(* IEC 61131-3 sources: plc-st-coding-agent/progress/evidence/f14_v6_public_pilot_20261112/jobs/custom_minimax-m27 (part 2) *)

(* ---- public-medium-03.candidate_02.st ---- *)
FUNCTION_BLOCK FB_MovingAverage
VAR_INPUT
    cyclicExecution : BOOL;
    trigger         : BOOL;
    value           : LREAL;
    windowSize      : INT;
    reset           : BOOL;
END_VAR

VAR_OUTPUT
    average           : LREAL;
    windowSizeReached : BOOL;
    error             : BOOL;
    status            : WORD;
END_VAR

VAR
    dataBuffer       : ARRAY[1..100] OF LREAL;
    currentIndex     : INT := 0;
    sampleCount      : INT := 0;
    sum              : LREAL := 0.0;
    tmp_lastTrigger  : BOOL := FALSE;
    tmp_newSample    : BOOL := FALSE;
    tmp_effectiveWin : INT := 0;
END_VAR

(*
ENGINEERING_CONTRACT
===================
Operation Modes:
- cyclicExecution=TRUE: Update every scan cycle; trigger ignored (PUB002)
- cyclicExecution=FALSE: Rising edge on trigger updates average (PUB003)
- reset=TRUE: Clear all state, outputs to default, status=SUCCESS (PUB004)

Output Retention Policy:
| Output             | Activation         | Retention    | Reset by reset=TRUE |
|--------------------|--------------------|--------------|---------------------|
| average            | Each valid sample  | Hold last    | Yes (→0.0)          |
| windowSizeReached  | sampleCount>=winSz | Hold TRUE    | Yes (→FALSE)        |
| error              | windowSize<1 or >100| Hold TRUE   | Yes (→FALSE)        |
| status             | Per validation     | Hold code    | Yes (→SUCCESS)      |

Boundary Conditions:
- windowSize<1 OR >100 → error=TRUE, status=16#8200, skip processing (PUB004, PUB007)
- reset asserted → immediate clear, no processing (PUB004)
- Empty window (sampleCount=0) → average=0.0 (division-safe)
- Circular buffer wraps at windowSize, never exceeds 100 elements

Same-Scan Priority:
1. reset check (highest)
2. windowSize validation
3. trigger rising-edge detection
4. cyclicExecution evaluation
5. sample insertion / buffer rotation
6. average recalculation

Units: LREAL for all arithmetic (PUB001). windowSize in slots [1..100].
*)

(* CONTRACT_RULES
[
  {"kind": "hold_until_reset", "output": "windowSizeReached", "set_input": null, "reset_input": "reset"},
  {"kind": "hold_until_reset", "output": "error", "set_input": null, "reset_input": "reset"},
  {"kind": "hold_until_reset", "output": "status", "set_input": null, "reset_input": "reset"}
]
*)

    // Reset: clear all state and outputs
    IF reset THEN
        currentIndex      := 0;
        sampleCount       := 0;
        sum               := 0.0;
        average           := 0.0;
        windowSizeReached := FALSE;
        error             := FALSE;
        status            := 16#0000;
        tmp_lastTrigger   := FALSE;
        tmp_newSample     := FALSE;
        tmp_effectiveWin  := 0;
        RETURN;
    END_IF;

    // Validate window size (PUB007)
    IF windowSize < 1 OR windowSize > 100 THEN
        error  := TRUE;
        status := 16#8200;
        RETURN;
    END_IF;

    // No validation error; set success status (PUB006)
    error  := FALSE;
    status := 16#0000;

    // Determine if a new sample should be processed (PUB002, PUB003)
    tmp_newSample := FALSE;
    IF cyclicExecution THEN
        tmp_newSample := TRUE;
    ELSIF trigger AND NOT tmp_lastTrigger THEN
        tmp_newSample := TRUE;
    END_IF;
    tmp_lastTrigger := trigger;

    // Process new data point if triggered (PUB001)
    IF tmp_newSample THEN
        // Clamp effective window to array upper bound (100)
        tmp_effectiveWin := windowSize;
        IF tmp_effectiveWin > 100 THEN
            tmp_effectiveWin := 100;
        END_IF;

        IF sampleCount < tmp_effectiveWin THEN
            // Window not yet full: append new value
            sampleCount := sampleCount + 1;
            dataBuffer[sampleCount] := value;
            sum := sum + value;
        ELSE
            // Window full: rotate out oldest value using circular buffer
            currentIndex := (currentIndex MOD tmp_effectiveWin) + 1;
            sum := sum - dataBuffer[currentIndex] + value;
            dataBuffer[currentIndex] := value;
        END_IF;
    END_IF;

    // Calculate moving arithmetic mean (PUB001)
    IF sampleCount > 0 THEN
        average := sum / TO_LREAL(sampleCount);
    ELSE
        average := 0.0;
    END_IF;

    // Indicate whether maximum window width has been reached (PUB001)
    tmp_effectiveWin := windowSize;
    IF tmp_effectiveWin > 100 THEN
        tmp_effectiveWin := 100;
    END_IF;
    windowSizeReached := (sampleCount >= tmp_effectiveWin);

END_FUNCTION_BLOCK

(* ---- public-medium-03.candidate_03.st ---- *)
FUNCTION_BLOCK FB_MovingAverage
VAR_INPUT
    cyclicExecution : BOOL;
    trigger         : BOOL;
    value           : LREAL;
    windowSize      : INT;
    reset           : BOOL;
END_VAR

VAR_OUTPUT
    average           : LREAL;
    windowSizeReached : BOOL;
    error             : BOOL;
    status            : WORD;
END_VAR

VAR
    dataBuffer       : ARRAY[1..100] OF LREAL;
    sampleCount      : INT := 0;
    sum              : LREAL := 0.0;
    tmp_lastTrigger  : BOOL := FALSE;
    tmp_effectiveWin : INT := 0;
END_VAR

(*
ENGINEERING_CONTRACT
===================
Operation Modes:
- cyclicExecution=TRUE: Update every scan cycle; trigger ignored (PUB002)
- cyclicExecution=FALSE: Rising edge on trigger updates average (PUB003)
- reset=TRUE: Clear all state, outputs to default, status=SUCCESS (PUB004)

Output Retention Policy:
| Output             | Activation         | Retention    | Reset by reset=TRUE |
|--------------------|--------------------|--------------|---------------------|
| average            | Each valid sample  | Hold last    | Yes (→0.0)          |
| windowSizeReached  | sampleCount>=winSz | Hold TRUE    | Yes (→FALSE)        |
| error              | windowSize<1 or >100| Hold TRUE   | Yes (→FALSE)        |
| status             | Per validation     | Hold code    | Yes (→SUCCESS)      |

Boundary Conditions:
- windowSize<1 OR >100 → error=TRUE, status=16#8200, skip processing (PUB004, PUB007)
- reset asserted → immediate clear, no processing (PUB004)
- Empty window (sampleCount=0) → average=0.0 (division-safe)
- Circular buffer wraps at windowSize, never exceeds 100 elements

Same-Scan Priority:
1. reset check (highest)
2. windowSize validation
3. trigger rising-edge detection
4. cyclicExecution evaluation
5. sample insertion / buffer rotation
6. average recalculation

Units: LREAL for all arithmetic (PUB001). windowSize in slots [1..100].
*)

(* CONTRACT_RULES
[
  {"kind": "hold_until_reset", "output": "windowSizeReached", "set_input": null, "reset_input": "reset"},
  {"kind": "hold_until_reset", "output": "error", "set_input": null, "reset_input": "reset"},
  {"kind": "hold_until_reset", "output": "status", "set_input": null, "reset_input": "reset"}
]
*)

    // Reset: clear all state and outputs
    IF reset THEN
        sampleCount       := 0;
        sum               := 0.0;
        average           := 0.0;
        windowSizeReached := FALSE;
        error             := FALSE;
        status            := 16#0000;
        tmp_lastTrigger   := FALSE;
        tmp_effectiveWin  := 0;
        RETURN;
    END_IF;

    // Validate window size (PUB007)
    IF windowSize < 1 OR windowSize > 100 THEN
        error  := TRUE;
        status := 16#8200;
        RETURN;
    END_IF;

    // No validation error; set success status (PUB006)
    error  := FALSE;
    status := 16#0000;

    // Clamp effective window to array upper bound (100)
    tmp_effectiveWin := windowSize;
    IF tmp_effectiveWin > 100 THEN
        tmp_effectiveWin := 100;
    END_IF;

    // Determine if a new sample should be processed (PUB002, PUB003)
    IF cyclicExecution OR (trigger AND NOT tmp_lastTrigger) THEN
        // Process new data point (PUB001)
        IF sampleCount < tmp_effectiveWin THEN
            // Window not yet full: append new value
            sampleCount := sampleCount + 1;
            dataBuffer[sampleCount] := value;
            sum := sum + value;
        ELSE
            // Window full: rotate out oldest value
            // Shift all elements down by one position
            sum := sum - dataBuffer[1];
            FOR i := 1 TO tmp_effectiveWin - 1 DO
                dataBuffer[i] := dataBuffer[i + 1];
            END_FOR;
            dataBuffer[tmp_effectiveWin] := value;
            sum := sum + value;
        END_IF;
    END_IF;

    // Update trigger state for edge detection
    tmp_lastTrigger := trigger;

    // Calculate moving arithmetic mean (PUB001)
    IF sampleCount > 0 THEN
        average := sum / TO_LREAL(sampleCount);
    ELSE
        average := 0.0;
    END_IF;

    // Indicate whether maximum window width has been reached (PUB001)
    windowSizeReached := (sampleCount >= tmp_effectiveWin);

END_FUNCTION_BLOCK

(* ---- public-medium-03.candidate_04.st ---- *)
FUNCTION_BLOCK FB_MovingAverage
VAR_INPUT
    cyclicExecution : BOOL;
    trigger         : BOOL;
    value           : LREAL;
    windowSize      : INT;
    reset           : BOOL;
END_VAR

VAR_OUTPUT
    average           : LREAL;
    windowSizeReached : BOOL;
    error             : BOOL;
    status            : WORD;
END_VAR

VAR
    dataBuffer         : ARRAY[1..100] OF LREAL;
    currentIndex       : INT := 0;
    sampleCount        : INT := 0;
    sum                : LREAL := 0.0;
    tmp_lastTrigger    : BOOL := FALSE;
    tmp_newSample      : BOOL := FALSE;
    tmp_effectiveWin   : INT := 0;
    tmp_winSizeChanged : BOOL := FALSE;
    tmp_prevWinSize    : INT := 0;
    tmp_startIdx       : INT := 0;
    tmp_i              : INT := 0;
    tmp_newSum         : LREAL := 0.0;
END_VAR

(*
ENGINEERING_CONTRACT
===================
Operation Modes:
- cyclicExecution=TRUE: Update every scan cycle; trigger ignored (PUB002)
- cyclicExecution=FALSE: Rising edge on trigger updates average (PUB003)
- reset=TRUE: Clear all state, outputs to default, status=SUCCESS (PUB004)

Output Retention Policy:
| Output             | Activation         | Retention    | Reset by reset=TRUE |
|--------------------|--------------------|--------------|---------------------|
| average            | Each valid sample  | Hold last    | Yes (→0.0)          |
| windowSizeReached  | sampleCount>=winSz | Hold TRUE    | Yes (→FALSE)        |
| error              | windowSize<1 or >100| Hold TRUE   | Yes (→FALSE)        |
| status             | Per validation     | Hold code    | Yes (→SUCCESS)      |

Boundary Conditions:
- windowSize<1 OR >100 → error=TRUE, status=16#8200, skip processing (PUB004, PUB007)
- reset asserted → immediate clear, no processing (PUB004)
- Empty window (sampleCount=0) → average=0.0 (division-safe)
- Circular buffer wraps at windowSize, never exceeds 100 elements
- windowSize change → prune buffer to contain only most recent windowSize samples

Same-Scan Priority:
1. reset check (highest)
2. windowSize validation (set error=TRUE if invalid, return)
3. windowSize change detection → prune buffer
4. trigger rising-edge detection
5. cyclicExecution evaluation
6. sample insertion / buffer rotation
7. average recalculation

Units: LREAL for all arithmetic (PUB001). windowSize in slots [1..100].
*)

(* CONTRACT_RULES
[
  {"kind": "hold_until_reset", "output": "windowSizeReached", "set_input": null, "reset_input": "reset"},
  {"kind": "hold_until_reset", "output": "error", "set_input": null, "reset_input": "reset"},
  {"kind": "hold_until_reset", "output": "status", "set_input": null, "reset_input": "reset"}
]
*)

    // Reset: clear all state and outputs
    IF reset THEN
        currentIndex      := 0;
        sampleCount       := 0;
        sum               := 0.0;
        average           := 0.0;
        windowSizeReached := FALSE;
        error             := FALSE;
        status            := 16#0000;
        tmp_lastTrigger   := FALSE;
        tmp_newSample     := FALSE;
        tmp_effectiveWin  := 0;
        tmp_winSizeChanged := FALSE;
        tmp_prevWinSize   := 0;
        tmp_startIdx      := 0;
        tmp_i             := 0;
        tmp_newSum        := 0.0;
        RETURN;
    END_IF;

    // Clamp effective window to array upper bound for validation
    tmp_effectiveWin := windowSize;
    IF tmp_effectiveWin > 100 THEN
        tmp_effectiveWin := 100;
    END_IF;

    // Validate window size (PUB007)
    // Only clear error AFTER validation passes, so invalid sizes preserve error state
    IF windowSize < 1 OR windowSize > 100 THEN
        error  := TRUE;
        status := 16#8200;
        RETURN;
    END_IF;

    // Valid windowSize: clear error and set success status (PUB006)
    error  := FALSE;
    status := 16#0000;

    // Detect windowSize change and prune buffer if needed
    tmp_winSizeChanged := (tmp_prevWinSize <> 0) AND (tmp_prevWinSize <> windowSize);
    IF tmp_winSizeChanged AND sampleCount > 0 THEN
        // Prune buffer to contain only most recent windowSize samples
        tmp_effectiveWin := windowSize;
        IF tmp_effectiveWin > 100 THEN
            tmp_effectiveWin := 100;
        END_IF;

        IF sampleCount > tmp_effectiveWin THEN
            // Calculate start index for circular buffer (oldest sample to keep)
            // Most recent samples are at positions (currentIndex - k + 1) through currentIndex
            tmp_startIdx := ((currentIndex - tmp_effectiveWin) MOD 100) + 1;
            IF tmp_startIdx < 1 THEN
                tmp_startIdx := tmp_startIdx + 100;
            END_IF;

            // Copy most recent samples to front of buffer and recalculate sum
            tmp_newSum := 0.0;
            FOR tmp_i := 1 TO tmp_effectiveWin DO
                dataBuffer[tmp_i] := dataBuffer[tmp_startIdx + tmp_i - 1];
                tmp_newSum := tmp_newSum + dataBuffer[tmp_i];
            END_FOR;

            // Clear remaining buffer slots
            FOR tmp_i := tmp_effectiveWin + 1 TO 100 DO
                dataBuffer[tmp_i] := 0.0;
            END_FOR;

            sampleCount := tmp_effectiveWin;
            sum := tmp_newSum;
            currentIndex := tmp_effectiveWin;
        END_IF;
    END_IF;

    // Track current windowSize for next-cycle change detection
    tmp_prevWinSize := windowSize;

    // Determine if a new sample should be processed (PUB002, PUB003)
    tmp_newSample := FALSE;
    IF cyclicExecution THEN
        tmp_newSample := TRUE;
    ELSIF trigger AND NOT tmp_lastTrigger THEN
        tmp_newSample := TRUE;
    END_IF;
    tmp_lastTrigger := trigger;

    // Process new data point if triggered (PUB001)
    IF tmp_newSample THEN
        tmp_effectiveWin := windowSize;
        IF tmp_effectiveWin > 100 THEN
            tmp_effectiveWin := 100;
        END_IF;

        IF sampleCount < tmp_effectiveWin THEN
            // Buffer not yet full: append new value
            sampleCount := sampleCount + 1;
            currentIndex := sampleCount;
            dataBuffer[currentIndex] := value;
            sum := sum + value;
        ELSE
            // Buffer full: rotate out oldest value using circular buffer
            currentIndex := (currentIndex MOD tmp_effectiveWin) + 1;
            sum := sum - dataBuffer[currentIndex] + value;
            dataBuffer[currentIndex] := value;
        END_IF;
    END_IF;

    // Calculate moving arithmetic mean (PUB001)
    IF sampleCount > 0 THEN
        average := sum / TO_LREAL(sampleCount);
    ELSE
        average := 0.0;
    END_IF;

    // Indicate whether maximum window width has been reached (PUB001)
    tmp_effectiveWin := windowSize;
    IF tmp_effectiveWin > 100 THEN
        tmp_effectiveWin := 100;
    END_IF;
    windowSizeReached := (sampleCount >= tmp_effectiveWin);

END_FUNCTION_BLOCK

(* ---- public-medium-03.raw_candidate_01.st ---- *)
FUNCTION_BLOCK FB_MovingAverage
VAR_INPUT
    cyclicExecution : BOOL;
    trigger         : BOOL;
    value           : LREAL;
    windowSize      : INT;
    reset           : BOOL;
END_VAR

VAR_OUTPUT
    average           : LREAL;
    windowSizeReached : BOOL;
    error             : BOOL;
    status            : WORD;
END_VAR

VAR
    dataBuffer    : ARRAY[1..100] OF LREAL;
    currentIndex  : INT := 0;
    sampleCount   : INT := 0;
    sum           : LREAL := 0.0;
    tmp_lastTrigger : BOOL := FALSE;
END_VAR

(*
ENGINEERING_CONTRACT
===================
Operation Modes:
- cyclicExecution=TRUE: Update every scan cycle; trigger ignored (PUB002)
- cyclicExecution=FALSE: Rising edge on trigger updates average (PUB003)
- reset=TRUE: Clear all state, outputs to default, status=SUCCESS (PUB004)

Output Retention Policy:
| Output             | Activation         | Retention    | Reset by reset=TRUE |
|--------------------|--------------------|--------------|---------------------|
| average            | Each valid sample  | Hold last    | Yes (→0.0)          |
| windowSizeReached  | sampleCount>=winSz | Hold TRUE    | Yes (→FALSE)        |
| error              | windowSize<1 or >100| Hold TRUE   | Yes (→FALSE)        |
| status             | Per validation     | Hold code    | Yes (→SUCCESS)      |

Boundary Conditions:
- windowSize<1 OR >100 → error=TRUE, status=16#8200, skip processing (PUB004, PUB007)
- reset asserted → immediate clear, no processing (PUB004)
- Empty window (sampleCount=0) → average=0.0 (division-safe)
- Circular buffer wraps at windowSize, never exceeds 100 elements

Same-Scan Priority:
1. reset check (highest)
2. windowSize validation
3. trigger rising-edge detection
4. cyclicExecution evaluation
5. sample insertion / buffer rotation
6. average recalculation

Units: LREAL for all arithmetic (PUB001). windowSize in slots [1..100].
*)

(* CONTRACT_RULES
[
  {"kind": "hold_until_reset", "output": "windowSizeReached", "set_input": null, "reset_input": "reset"},
  {"kind": "hold_until_reset", "output": "error", "set_input": null, "reset_input": "reset"},
  {"kind": "hold_until_reset", "output": "status", "set_input": null, "reset_input": "reset"}
]
*)

    // Reset: clear all state and outputs
    IF reset THEN
        currentIndex     := 0;
        sampleCount      := 0;
        sum              := 0.0;
        average          := 0.0;
        windowSizeReached := FALSE;
        error            := FALSE;
        status           := 16#0000;
        tmp_lastTrigger  := FALSE;
        RETURN;
    END_IF

    // Validate window size (PUB007)
    IF windowSize < 1 OR windowSize > 100 THEN
        error  := TRUE;
        status := 16#8200;
        RETURN;
    END_IF

    // No validation error; set success status (PUB006)
    error  := FALSE;
    status := 16#0000;

    // Determine if a new sample should be processed (PUB002, PUB003)
    tmp_newSample := FALSE;
    IF cyclicExecution THEN
        tmp_newSample := TRUE;
    ELSIF trigger AND NOT tmp_lastTrigger THEN
        tmp_newSample := TRUE;
    END_IF
    tmp_lastTrigger := trigger;

    // Process new data point if triggered (PUB001)
    IF tmp_newSample THEN
        // Clamp effective window to array upper bound (100)
        tmp_effectiveWindow := windowSize;
        IF tmp_effectiveWindow > 100 THEN
            tmp_effectiveWindow := 100;
        END_IF

        IF sampleCount < tmp_effectiveWindow THEN
            // Window not yet full: append new value
            sampleCount := sampleCount + 1;
            dataBuffer[sampleCount] := value;
            sum := sum + value;
        ELSE
            // Window full: rotate out oldest value using circular buffer
            currentIndex := (currentIndex MOD tmp_effectiveWindow) + 1;
            sum := sum - dataBuffer[currentIndex] + value;
            dataBuffer[currentIndex] := value;
        END_IF
    END_IF

    // Calculate moving arithmetic mean (PUB001)
    IF sampleCount > 0 THEN
        average := sum / TO_LREAL(sampleCount);
    ELSE
        average := 0.0;
    END_IF

    // Indicate whether maximum window width has been reached (PUB001)
    tmp_effectiveWindow := windowSize;
    IF tmp_effectiveWindow > 100 THEN
        tmp_effectiveWindow := 100;
    END_IF;
    windowSizeReached := (sampleCount >= tmp_effectiveWindow);

END_FUNCTION_BLOCK

(* ---- public-medium-03.raw_candidate_02.st ---- *)
FUNCTION_BLOCK FB_MovingAverage
VAR_INPUT
    cyclicExecution : BOOL;
    trigger         : BOOL;
    value           : LREAL;
    windowSize      : INT;
    reset           : BOOL;
END_VAR

VAR_OUTPUT
    average           : LREAL;
    windowSizeReached : BOOL;
    error             : BOOL;
    status            : WORD;
END_VAR

VAR
    dataBuffer       : ARRAY[1..100] OF LREAL;
    currentIndex     : INT := 0;
    sampleCount      : INT := 0;
    sum              : LREAL := 0.0;
    tmp_lastTrigger  : BOOL := FALSE;
    tmp_newSample    : BOOL := FALSE;
    tmp_effectiveWin : INT := 0;
END_VAR

(*
ENGINEERING_CONTRACT
===================
Operation Modes:
- cyclicExecution=TRUE: Update every scan cycle; trigger ignored (PUB002)
- cyclicExecution=FALSE: Rising edge on trigger updates average (PUB003)
- reset=TRUE: Clear all state, outputs to default, status=SUCCESS (PUB004)

Output Retention Policy:
| Output             | Activation         | Retention    | Reset by reset=TRUE |
|--------------------|--------------------|--------------|---------------------|
| average            | Each valid sample  | Hold last    | Yes (→0.0)          |
| windowSizeReached  | sampleCount>=winSz | Hold TRUE    | Yes (→FALSE)        |
| error              | windowSize<1 or >100| Hold TRUE   | Yes (→FALSE)        |
| status             | Per validation     | Hold code    | Yes (→SUCCESS)      |

Boundary Conditions:
- windowSize<1 OR >100 → error=TRUE, status=16#8200, skip processing (PUB004, PUB007)
- reset asserted → immediate clear, no processing (PUB004)
- Empty window (sampleCount=0) → average=0.0 (division-safe)
- Circular buffer wraps at windowSize, never exceeds 100 elements

Same-Scan Priority:
1. reset check (highest)
2. windowSize validation
3. trigger rising-edge detection
4. cyclicExecution evaluation
5. sample insertion / buffer rotation
6. average recalculation

Units: LREAL for all arithmetic (PUB001). windowSize in slots [1..100].
*)

(* CONTRACT_RULES
[
  {"kind": "hold_until_reset", "output": "windowSizeReached", "set_input": null, "reset_input": "reset"},
  {"kind": "hold_until_reset", "output": "error", "set_input": null, "reset_input": "reset"},
  {"kind": "hold_until_reset", "output": "status", "set_input": null, "reset_input": "reset"}
]
*)

    // Reset: clear all state and outputs
    IF reset THEN
        currentIndex      := 0;
        sampleCount       := 0;
        sum               := 0.0;
        average           := 0.0;
        windowSizeReached := FALSE;
        error             := FALSE;
        status            := 16#0000;
        tmp_lastTrigger   := FALSE;
        tmp_newSample     := FALSE;
        tmp_effectiveWin  := 0;
        RETURN;
    END_IF;

    // Validate window size (PUB007)
    IF windowSize < 1 OR windowSize > 100 THEN
        error  := TRUE;
        status := 16#8200;
        RETURN;
    END_IF;

    // No validation error; set success status (PUB006)
    error  := FALSE;
    status := 16#0000;

    // Determine if a new sample should be processed (PUB002, PUB003)
    tmp_newSample := FALSE;
    IF cyclicExecution THEN
        tmp_newSample := TRUE;
    ELSIF trigger AND NOT tmp_lastTrigger THEN
        tmp_newSample := TRUE;
    END_IF;
    tmp_lastTrigger := trigger;

    // Process new data point if triggered (PUB001)
    IF tmp_newSample THEN
        // Clamp effective window to array upper bound (100)
        tmp_effectiveWin := windowSize;
        IF tmp_effectiveWin > 100 THEN
            tmp_effectiveWin := 100;
        END_IF;

        IF sampleCount < tmp_effectiveWin THEN
            // Window not yet full: append new value
            sampleCount := sampleCount + 1;
            dataBuffer[sampleCount] := value;
            sum := sum + value;
        ELSE
            // Window full: rotate out oldest value using circular buffer
            currentIndex := (currentIndex MOD tmp_effectiveWin) + 1;
            sum := sum - dataBuffer[currentIndex] + value;
            dataBuffer[currentIndex] := value;
        END_IF;
    END_IF;

    // Calculate moving arithmetic mean (PUB001)
    IF sampleCount > 0 THEN
        average := sum / TO_LREAL(sampleCount);
    ELSE
        average := 0.0;
    END_IF;

    // Indicate whether maximum window width has been reached (PUB001)
    tmp_effectiveWin := windowSize;
    IF tmp_effectiveWin > 100 THEN
        tmp_effectiveWin := 100;
    END_IF;
    windowSizeReached := (sampleCount >= tmp_effectiveWin);

END_FUNCTION_BLOCK

(* ---- public-medium-03.raw_candidate_03.st ---- *)
FUNCTION_BLOCK FB_MovingAverage
VAR_INPUT
    cyclicExecution : BOOL;
    trigger         : BOOL;
    value           : LREAL;
    windowSize      : INT;
    reset           : BOOL;
END_VAR

VAR_OUTPUT
    average           : LREAL;
    windowSizeReached : BOOL;
    error             : BOOL;
    status            : WORD;
END_VAR

VAR
    dataBuffer       : ARRAY[1..100] OF LREAL;
    sampleCount      : INT := 0;
    sum              : LREAL := 0.0;
    tmp_lastTrigger  : BOOL := FALSE;
    tmp_effectiveWin : INT := 0;
END_VAR

(*
ENGINEERING_CONTRACT
===================
Operation Modes:
- cyclicExecution=TRUE: Update every scan cycle; trigger ignored (PUB002)
- cyclicExecution=FALSE: Rising edge on trigger updates average (PUB003)
- reset=TRUE: Clear all state, outputs to default, status=SUCCESS (PUB004)

Output Retention Policy:
| Output             | Activation         | Retention    | Reset by reset=TRUE |
|--------------------|--------------------|--------------|---------------------|
| average            | Each valid sample  | Hold last    | Yes (→0.0)          |
| windowSizeReached  | sampleCount>=winSz | Hold TRUE    | Yes (→FALSE)        |
| error              | windowSize<1 or >100| Hold TRUE   | Yes (→FALSE)        |
| status             | Per validation     | Hold code    | Yes (→SUCCESS)      |

Boundary Conditions:
- windowSize<1 OR >100 → error=TRUE, status=16#8200, skip processing (PUB004, PUB007)
- reset asserted → immediate clear, no processing (PUB004)
- Empty window (sampleCount=0) → average=0.0 (division-safe)
- Circular buffer wraps at windowSize, never exceeds 100 elements

Same-Scan Priority:
1. reset check (highest)
2. windowSize validation
3. trigger rising-edge detection
4. cyclicExecution evaluation
5. sample insertion / buffer rotation
6. average recalculation

Units: LREAL for all arithmetic (PUB001). windowSize in slots [1..100].
*)

(* CONTRACT_RULES
[
  {"kind": "hold_until_reset", "output": "windowSizeReached", "set_input": null, "reset_input": "reset"},
  {"kind": "hold_until_reset", "output": "error", "set_input": null, "reset_input": "reset"},
  {"kind": "hold_until_reset", "output": "status", "set_input": null, "reset_input": "reset"}
]
*)

    // Reset: clear all state and outputs
    IF reset THEN
        sampleCount       := 0;
        sum               := 0.0;
        average           := 0.0;
        windowSizeReached := FALSE;
        error             := FALSE;
        status            := 16#0000;
        tmp_lastTrigger   := FALSE;
        tmp_effectiveWin  := 0;
        RETURN;
    END_IF;

    // Validate window size (PUB007)
    IF windowSize < 1 OR windowSize > 100 THEN
        error  := TRUE;
        status := 16#8200;
        RETURN;
    END_IF;

    // No validation error; set success status (PUB006)
    error  := FALSE;
    status := 16#0000;

    // Clamp effective window to array upper bound (100)
    tmp_effectiveWin := windowSize;
    IF tmp_effectiveWin > 100 THEN
        tmp_effectiveWin := 100;
    END_IF;

    // Determine if a new sample should be processed (PUB002, PUB003)
    IF cyclicExecution OR (trigger AND NOT tmp_lastTrigger) THEN
        // Process new data point (PUB001)
        IF sampleCount < tmp_effectiveWin THEN
            // Window not yet full: append new value
            sampleCount := sampleCount + 1;
            dataBuffer[sampleCount] := value;
            sum := sum + value;
        ELSE
            // Window full: rotate out oldest value
            // Shift all elements down by one position
            sum := sum - dataBuffer[1];
            FOR i := 1 TO tmp_effectiveWin - 1 DO
                dataBuffer[i] := dataBuffer[i + 1];
            END_FOR;
            dataBuffer[tmp_effectiveWin] := value;
            sum := sum + value;
        END_IF;
    END_IF;

    // Update trigger state for edge detection
    tmp_lastTrigger := trigger;

    // Calculate moving arithmetic mean (PUB001)
    IF sampleCount > 0 THEN
        average := sum / TO_LREAL(sampleCount);
    ELSE
        average := 0.0;
    END_IF;

    // Indicate whether maximum window width has been reached (PUB001)
    windowSizeReached := (sampleCount >= tmp_effectiveWin);

END_FUNCTION_BLOCK

(* ---- public-medium-03.raw_candidate_04.st ---- *)
FUNCTION_BLOCK FB_MovingAverage
VAR_INPUT
    cyclicExecution : BOOL;
    trigger         : BOOL;
    value           : LREAL;
    windowSize      : INT;
    reset           : BOOL;
END_VAR

VAR_OUTPUT
    average           : LREAL;
    windowSizeReached : BOOL;
    error             : BOOL;
    status            : WORD;
END_VAR

VAR
    dataBuffer         : ARRAY[1..100] OF LREAL;
    currentIndex       : INT := 0;
    sampleCount        : INT := 0;
    sum                : LREAL := 0.0;
    tmp_lastTrigger    : BOOL := FALSE;
    tmp_newSample      : BOOL := FALSE;
    tmp_effectiveWin   : INT := 0;
    tmp_winSizeChanged : BOOL := FALSE;
    tmp_prevWinSize    : INT := 0;
    tmp_startIdx       : INT := 0;
    tmp_i              : INT := 0;
    tmp_newSum         : LREAL := 0.0;
END_VAR

(*
ENGINEERING_CONTRACT
===================
Operation Modes:
- cyclicExecution=TRUE: Update every scan cycle; trigger ignored (PUB002)
- cyclicExecution=FALSE: Rising edge on trigger updates average (PUB003)
- reset=TRUE: Clear all state, outputs to default, status=SUCCESS (PUB004)

Output Retention Policy:
| Output             | Activation         | Retention    | Reset by reset=TRUE |
|--------------------|--------------------|--------------|---------------------|
| average            | Each valid sample  | Hold last    | Yes (→0.0)          |
| windowSizeReached  | sampleCount>=winSz | Hold TRUE    | Yes (→FALSE)        |
| error              | windowSize<1 or >100| Hold TRUE   | Yes (→FALSE)        |
| status             | Per validation     | Hold code    | Yes (→SUCCESS)      |

Boundary Conditions:
- windowSize<1 OR >100 → error=TRUE, status=16#8200, skip processing (PUB004, PUB007)
- reset asserted → immediate clear, no processing (PUB004)
- Empty window (sampleCount=0) → average=0.0 (division-safe)
- Circular buffer wraps at windowSize, never exceeds 100 elements
- windowSize change → prune buffer to contain only most recent windowSize samples

Same-Scan Priority:
1. reset check (highest)
2. windowSize validation (set error=TRUE if invalid, return)
3. windowSize change detection → prune buffer
4. trigger rising-edge detection
5. cyclicExecution evaluation
6. sample insertion / buffer rotation
7. average recalculation

Units: LREAL for all arithmetic (PUB001). windowSize in slots [1..100].
*)

(* CONTRACT_RULES
[
  {"kind": "hold_until_reset", "output": "windowSizeReached", "set_input": null, "reset_input": "reset"},
  {"kind": "hold_until_reset", "output": "error", "set_input": null, "reset_input": "reset"},
  {"kind": "hold_until_reset", "output": "status", "set_input": null, "reset_input": "reset"}
]
*)

    // Reset: clear all state and outputs
    IF reset THEN
        currentIndex      := 0;
        sampleCount       := 0;
        sum               := 0.0;
        average           := 0.0;
        windowSizeReached := FALSE;
        error             := FALSE;
        status            := 16#0000;
        tmp_lastTrigger   := FALSE;
        tmp_newSample     := FALSE;
        tmp_effectiveWin  := 0;
        tmp_winSizeChanged := FALSE;
        tmp_prevWinSize   := 0;
        tmp_startIdx      := 0;
        tmp_i             := 0;
        tmp_newSum        := 0.0;
        RETURN;
    END_IF;

    // Clamp effective window to array upper bound for validation
    tmp_effectiveWin := windowSize;
    IF tmp_effectiveWin > 100 THEN
        tmp_effectiveWin := 100;
    END_IF;

    // Validate window size (PUB007)
    // Only clear error AFTER validation passes, so invalid sizes preserve error state
    IF windowSize < 1 OR windowSize > 100 THEN
        error  := TRUE;
        status := 16#8200;
        RETURN;
    END_IF;

    // Valid windowSize: clear error and set success status (PUB006)
    error  := FALSE;
    status := 16#0000;

    // Detect windowSize change and prune buffer if needed
    tmp_winSizeChanged := (tmp_prevWinSize <> 0) AND (tmp_prevWinSize <> windowSize);
    IF tmp_winSizeChanged AND sampleCount > 0 THEN
        // Prune buffer to contain only most recent windowSize samples
        tmp_effectiveWin := windowSize;
        IF tmp_effectiveWin > 100 THEN
            tmp_effectiveWin := 100;
        END_IF;

        IF sampleCount > tmp_effectiveWin THEN
            // Calculate start index for circular buffer (oldest sample to keep)
            // Most recent samples are at positions (currentIndex - k + 1) through currentIndex
            tmp_startIdx := ((currentIndex - tmp_effectiveWin) MOD 100) + 1;
            IF tmp_startIdx < 1 THEN
                tmp_startIdx := tmp_startIdx + 100;
            END_IF;

            // Copy most recent samples to front of buffer and recalculate sum
            tmp_newSum := 0.0;
            FOR tmp_i := 1 TO tmp_effectiveWin DO
                dataBuffer[tmp_i] := dataBuffer[tmp_startIdx + tmp_i - 1];
                tmp_newSum := tmp_newSum + dataBuffer[tmp_i];
            END_FOR;

            // Clear remaining buffer slots
            FOR tmp_i := tmp_effectiveWin + 1 TO 100 DO
                dataBuffer[tmp_i] := 0.0;
            END_FOR;

            sampleCount := tmp_effectiveWin;
            sum := tmp_newSum;
            currentIndex := tmp_effectiveWin;
        END_IF;
    END_IF;

    // Track current windowSize for next-cycle change detection
    tmp_prevWinSize := windowSize;

    // Determine if a new sample should be processed (PUB002, PUB003)
    tmp_newSample := FALSE;
    IF cyclicExecution THEN
        tmp_newSample := TRUE;
    ELSIF trigger AND NOT tmp_lastTrigger THEN
        tmp_newSample := TRUE;
    END_IF;
    tmp_lastTrigger := trigger;

    // Process new data point if triggered (PUB001)
    IF tmp_newSample THEN
        tmp_effectiveWin := windowSize;
        IF tmp_effectiveWin > 100 THEN
            tmp_effectiveWin := 100;
        END_IF;

        IF sampleCount < tmp_effectiveWin THEN
            // Buffer not yet full: append new value
            sampleCount := sampleCount + 1;
            currentIndex := sampleCount;
            dataBuffer[currentIndex] := value;
            sum := sum + value;
        ELSE
            // Buffer full: rotate out oldest value using circular buffer
            currentIndex := (currentIndex MOD tmp_effectiveWin) + 1;
            sum := sum - dataBuffer[currentIndex] + value;
            dataBuffer[currentIndex] := value;
        END_IF;
    END_IF;

    // Calculate moving arithmetic mean (PUB001)
    IF sampleCount > 0 THEN
        average := sum / TO_LREAL(sampleCount);
    ELSE
        average := 0.0;
    END_IF;

    // Indicate whether maximum window width has been reached (PUB001)
    tmp_effectiveWin := windowSize;
    IF tmp_effectiveWin > 100 THEN
        tmp_effectiveWin := 100;
    END_IF;
    windowSizeReached := (sampleCount >= tmp_effectiveWin);

END_FUNCTION_BLOCK

(* ---- public-medium-04.candidate_01.st ---- *)
FUNCTION_BLOCK FBTemperatureControl
VAR_INPUT
    TemperatureSensorInput : REAL;
    SetTemperature         : REAL;
END_VAR
VAR_OUTPUT
    CurrentTemperature : REAL;
    SetTempDisplay     : REAL;
    HeaterStatus       : BOOL;
    OverheatProtection : BOOL;
    HeaterOutput       : BOOL := FALSE;
END_VAR
VAR
    tonHeaterRuntime   : TON;
    tonOverheatCooldown: TON;
    tmpSensorFault     : BOOL;
    tmpHeaterShouldBeOn: BOOL;
END_VAR

(* ENGINEERING_CONTRACT:
 * | State/Output       | Activation                          | Retention           | Reset/Deactivation                                      | Same-scan Priority     | Units/Boundaries   |
 * |--------------------|-------------------------------------|---------------------|---------------------------------------------------------|------------------------|--------------------|
 * | HeaterOutput       | Temp < SetTemp AND no fault AND no overheat | Held per scan       | Temp >= SetTemp OR fault OR overheat triggered          | Overheat overrides     | BOOLEAN            |
 * | OverheatProtection | HeaterOutput TRUE for >= 5s continuous  | Held until 3s cooldown done | After 3s cooldown done AND heater would be OFF | Timer-driven, latch    | BOOLEAN            |
 * | SensorFault        | Temp < 0 OR Temp > 100              | N/A (implicit)      | When temp returns to valid range                        | Implicit               | BOOLEAN (derived)  |
 * | HeaterStatus       | HeaterOutput = TRUE                 | Same as HeaterOutput | Same as HeaterOutput                                   | Display only           | BOOLEAN            |
 * | CurrentTemperature | Always updated                      | Per scan            | N/A                                                     | Always active          | REAL, 0-100 valid  |
 *)

(* CONTRACT_RULES [{"kind":"hold_until_reset","output":"HeaterOutput","set_input":"OverheatProtection","reset_input":null}] *)

tmpSensorFault := (TemperatureSensorInput < 0.0) OR (TemperatureSensorInput > 100.0);

tmpHeaterShouldBeOn := (TemperatureSensorInput < SetTemperature) AND (NOT tmpSensorFault) AND (NOT OverheatProtection);

IF OverheatProtection THEN
    tonHeaterRuntime(IN := FALSE, PT := T#5S);
    tonOverheatCooldown(IN := TRUE, PT := T#3S);
    IF tonOverheatCooldown.Q THEN
        OverheatProtection := FALSE;
        tonOverheatCooldown(IN := FALSE, PT := T#3S);
    END_IF;
ELSIF tmpHeaterShouldBeOn THEN
    tonOverheatCooldown(IN := FALSE, PT := T#3S);
    tonHeaterRuntime(IN := TRUE, PT := T#5S);
    IF tonHeaterRuntime.Q THEN
        OverheatProtection := TRUE;
        HeaterOutput := FALSE;
    ELSE
        HeaterOutput := TRUE;
    END_IF;
ELSE
    tonHeaterRuntime(IN := FALSE, PT := T#5S);
    tonOverheatCooldown(IN := FALSE, PT := T#3S);
    HeaterOutput := FALSE;
END_IF;

CurrentTemperature := TemperatureSensorInput;
SetTempDisplay     := SetTemperature;
HeaterStatus       := HeaterOutput;

END_FUNCTION_BLOCK

(* ---- public-medium-04.candidate_02.st ---- *)
FUNCTION_BLOCK FBTemperatureControl
VAR_INPUT
    TemperatureSensorInput : REAL;
    SetTemperature         : REAL;
END_VAR
VAR_OUTPUT
    CurrentTemperature : REAL;
    SetTempDisplay     : REAL;
    HeaterStatus       : BOOL;
    OverheatProtection : BOOL;
    HeaterOutput       : BOOL := FALSE;
END_VAR
VAR
    tonHeaterRuntime   : TON;
    tonOverheatCooldown: TON;
    tmpSensorFault     : BOOL;
END_VAR

(* ENGINEERING_CONTRACT:
 * | State/Output       | Activation                          | Retention           | Reset/Deactivation                                      | Same-scan Priority     | Units/Boundaries   |
 * |--------------------|-------------------------------------|---------------------|---------------------------------------------------------|------------------------|--------------------|
 * | HeaterOutput       | Temp < SetTemp AND no fault AND no overheat | Held per scan       | Temp >= SetTemp OR fault OR overheat triggered          | Overheat overrides     | BOOLEAN            |
 * | OverheatProtection | HeaterOutput TRUE for >= 5s continuous  | Held until 3s cooldown done | After 3s cooldown done AND heater would be OFF | Timer-driven, latch    | BOOLEAN            |
 * | SensorFault        | Temp < 0 OR Temp > 100              | N/A (implicit)      | When temp returns to valid range                        | Implicit               | BOOLEAN (derived)  |
 * | HeaterStatus       | HeaterOutput = TRUE                 | Same as HeaterOutput | Same as HeaterOutput                                   | Display only           | BOOLEAN            |
 * | CurrentTemperature | Always updated                      | Per scan            | N/A                                                     | Always active          | REAL, 0-100 valid  |
 *)

(* CONTRACT_RULES [] *)

tmpSensorFault := (TemperatureSensorInput < 0.0) OR (TemperatureSensorInput > 100.0);

IF OverheatProtection THEN
    tonHeaterRuntime(IN := FALSE, PT := T#0S);
    tonOverheatCooldown(IN := TRUE, PT := T#3S);
    IF tonOverheatCooldown.Q THEN
        OverheatProtection := FALSE;
        tonOverheatCooldown(IN := FALSE, PT := T#0S);
    END_IF;
    HeaterOutput := FALSE;
ELSIF (TemperatureSensorInput < SetTemperature) AND (NOT tmpSensorFault) THEN
    tonOverheatCooldown(IN := FALSE, PT := T#0S);
    tonHeaterRuntime(IN := TRUE, PT := T#5S);
    IF tonHeaterRuntime.Q THEN
        OverheatProtection := TRUE;
        HeaterOutput := FALSE;
        tonHeaterRuntime(IN := FALSE, PT := T#0S);
    ELSE
        HeaterOutput := TRUE;
    END_IF;
ELSE
    tonHeaterRuntime(IN := FALSE, PT := T#0S);
    tonOverheatCooldown(IN := FALSE, PT := T#0S);
    HeaterOutput := FALSE;
END_IF;

CurrentTemperature := TemperatureSensorInput;
SetTempDisplay     := SetTemperature;
HeaterStatus       := HeaterOutput;

END_FUNCTION_BLOCK

(* ---- public-medium-04.candidate_03.st ---- *)
FUNCTION_BLOCK FBTemperatureControl
VAR_INPUT
    TemperatureSensorInput : REAL;
    SetTemperature         : REAL;
END_VAR
VAR_OUTPUT
    CurrentTemperature : REAL;
    SetTempDisplay     : REAL;
    HeaterStatus       : BOOL;
    OverheatProtection : BOOL;
    HeaterOutput       : BOOL := FALSE;
END_VAR
VAR
    tonOverheatCooldown : TON;
    tmpSensorFault      : BOOL;
    tmpHeaterShouldBeOn : BOOL;
    tmpHeaterOn         : BOOL;
    tmpRuntimeAccum     : LTIME;  // Track accumulated heating time
    tmpCooldownAccum    : LTIME;  // Track cooldown elapsed time
END_VAR

(* ENGINEERING_CONTRACT:
 * | State/Output       | Activation                          | Retention           | Reset/Deactivation                                      | Same-scan Priority     | Units/Boundaries   |
 * |--------------------|-------------------------------------|---------------------|---------------------------------------------------------|------------------------|--------------------|
 * | HeaterOutput       | Temp < SetTemp AND no fault AND no overheat | Held per scan   | Temp >= SetTemp OR fault OR overheat triggered          | Overheat overrides     | BOOLEAN            |
 * | OverheatProtection | Runtime >= 5s continuous heater ON  | Held until 3s cooldown done | After 3s cooldown done AND heater would be OFF | Timer-driven, latch    | BOOLEAN            |
 * | SensorFault        | Temp < 0 OR Temp > 100              | N/A (implicit)      | When temp returns to valid range                        | Implicit               | BOOLEAN (derived)  |
 * | HeaterStatus       | HeaterOutput = TRUE                 | Same as HeaterOutput | Same as HeaterOutput                                   | Display only           | BOOLEAN            |
 * | CurrentTemperature | Always updated                      | Per scan            | N/A                                                     | Always active          | REAL, 0-100 valid  |
 * | RuntimeAccum       | Increments when heater ON, no overheat | Per scan         | Reset when heater OFF OR overheat triggers             | Counter-based          | LTIME, max 5s      |
 * | CooldownAccum      | Increments when OverheatProtection TRUE | Per scan        | Reset when OverheatProtection clears                   | Counter-based          | LTIME, max 3s      |
 *)

(* CONTRACT_RULES [] *)

tmpSensorFault := (TemperatureSensorInput < 0.0) OR (TemperatureSensorInput > 100.0);

tmpHeaterOn := FALSE;

IF OverheatProtection THEN
    // Cooldown phase: heater stays off, track cooldown time
    tonOverheatCooldown(IN := TRUE, PT := T#3S);
    tmpCooldownAccum := tmpCooldownAccum + LTIME#1ms;  // Framework advances 1ms per call

    IF tonOverheatCooldown.Q THEN
        OverheatProtection := FALSE;
        tmpRuntimeAccum := LTIME#0ms;
        tonOverheatCooldown(IN := FALSE, PT := T#3S);
    END_IF;

ELSIF (NOT tmpSensorFault) AND (TemperatureSensorInput < SetTemperature) THEN
    // Normal heating: heater can be ON
    tonOverheatCooldown(IN := FALSE, PT := T#3S);

    tmpRuntimeAccum := tmpRuntimeAccum + LTIME#1ms;  // Framework advances 1ms per call

    IF tmpRuntimeAccum >= LTIME#5000ms THEN
        // Overheat threshold reached
        OverheatProtection := TRUE;
        HeaterOutput       := FALSE;
        tmpHeaterOn        := FALSE;
        tmpCooldownAccum   := LTIME#0ms;
    ELSE
        HeaterOutput := TRUE;
        tmpHeaterOn  := TRUE;
    END_IF;

ELSE
    // Temperature OK or sensor fault: heater OFF
    tonOverheatCooldown(IN := FALSE, PT := T#3S);
    HeaterOutput    := FALSE;
    tmpHeaterOn     := FALSE;
    tmpRuntimeAccum := LTIME#0ms;
END_IF;

CurrentTemperature := TemperatureSensorInput;
SetTempDisplay     := SetTemperature;
HeaterStatus       := tmpHeaterOn;

END_FUNCTION_BLOCK

(* ---- public-medium-04.candidate_04.st ---- *)
FUNCTION_BLOCK FBTemperatureControl
VAR_INPUT
    TemperatureSensorInput : REAL;
    SetTemperature         : REAL;
END_VAR
VAR_OUTPUT
    CurrentTemperature : REAL;
    SetTempDisplay     : REAL;
    HeaterStatus       : BOOL;
    OverheatProtection : BOOL := FALSE;
    HeaterOutput       : BOOL := FALSE;
END_VAR
VAR
    tonHeaterRuntime   : TON;
    tonOverheatCooldown: TON;
    tmpSensorFault     : BOOL;
    tmpHeaterShouldBeOn: BOOL;
    tmpHeaterLatchedOff: BOOL := FALSE;
END_VAR

(* ENGINEERING_CONTRACT:
 * | State/Output       | Activation                          | Retention           | Reset/Deactivation                                      | Same-scan Priority     | Units/Boundaries   |
 * |--------------------|-------------------------------------|---------------------|---------------------------------------------------------|------------------------|--------------------|
 * | HeaterOutput       | Temp < SetTemp AND no fault AND no overheat/latch | Held per scan       | Temp >= SetTemp OR fault OR overheat/latch triggered    | Overheat overrides     | BOOLEAN            |
 * | OverheatProtection | HeaterOutput TRUE for >= 5s continuous  | Held until 3s cooldown done | After 3s cooldown done AND heater would be OFF | Timer-driven, latch    | BOOLEAN            |
 * | HeaterLatchedOff   | OverheatProtection triggers          | Held indefinitely   | No reset defined; remains latched                       | Latch persists         | BOOLEAN            |
 * | SensorFault        | Temp < 0 OR Temp > 100              | N/A (implicit)      | When temp returns to valid range                        | Implicit               | BOOLEAN (derived)  |
 * | HeaterStatus       | HeaterOutput = TRUE                 | Same as HeaterOutput | Same as HeaterOutput                                   | Display only           | BOOLEAN            |
 * | CurrentTemperature | Always updated                      | Per scan            | N/A                                                     | Always active          | REAL, 0-100 valid  |
 *)

(* CONTRACT_RULES [{"kind":"hold_until_reset","output":"HeaterOutput","set_input":"OverheatProtection","reset_input":null}] *)

tmpSensorFault := (TemperatureSensorInput < 0.0) OR (TemperatureSensorInput > 100.0);

IF OverheatProtection THEN
    tonHeaterRuntime(IN := FALSE, PT := T#5S);
    tonOverheatCooldown(IN := TRUE, PT := T#3S);
    IF tonOverheatCooldown.Q THEN
        OverheatProtection := FALSE;
        tmpHeaterLatchedOff := TRUE;
        tonOverheatCooldown(IN := FALSE, PT := T#3S);
        tonHeaterRuntime(IN := FALSE, PT := T#5S);
    END_IF;
    HeaterOutput := FALSE;
ELSIF tmpSensorFault THEN
    tonHeaterRuntime(IN := FALSE, PT := T#5S);
    tonOverheatCooldown(IN := FALSE, PT := T#3S);
    HeaterOutput := FALSE;
    tmpHeaterLatchedOff := FALSE;
ELSE
    tonOverheatCooldown(IN := FALSE, PT := T#3S);
    tmpHeaterShouldBeOn := (TemperatureSensorInput < SetTemperature) AND (NOT tmpHeaterLatchedOff);
    tonHeaterRuntime(IN := tmpHeaterShouldBeOn, PT := T#5S);
    IF tonHeaterRuntime.Q THEN
        OverheatProtection := TRUE;
        tmpHeaterLatchedOff := TRUE;
        HeaterOutput := FALSE;
    ELSIF tmpHeaterShouldBeOn THEN
        HeaterOutput := TRUE;
    ELSE
        HeaterOutput := FALSE;
        tmpHeaterLatchedOff := FALSE;
    END_IF;
END_IF;

CurrentTemperature := TemperatureSensorInput;
SetTempDisplay     := SetTemperature;
HeaterStatus       := HeaterOutput;

END_FUNCTION_BLOCK

(* ---- public-medium-04.raw_candidate_01.st ---- *)
FUNCTION_BLOCK FBTemperatureControl
VAR_INPUT
    TemperatureSensorInput : REAL;
    SetTemperature         : REAL;
END_VAR
VAR_OUTPUT
    CurrentTemperature : REAL;
    SetTempDisplay     : REAL;
    HeaterStatus       : BOOL;
    OverheatProtection : BOOL;
    HeaterOutput       : BOOL := FALSE;
END_VAR
VAR
    tonHeaterRuntime   : TON;
    tonOverheatCooldown: TON;
    tmpSensorFault     : BOOL;
    tmpHeaterShouldBeOn: BOOL;
END_VAR

(* ENGINEERING_CONTRACT:
 * | State/Output       | Activation                          | Retention           | Reset/Deactivation                                      | Same-scan Priority     | Units/Boundaries   |
 * |--------------------|-------------------------------------|---------------------|---------------------------------------------------------|------------------------|--------------------|
 * | HeaterOutput       | Temp < SetTemp AND no fault AND no overheat | Held per scan       | Temp >= SetTemp OR fault OR overheat triggered          | Overheat overrides     | BOOLEAN            |
 * | OverheatProtection | HeaterOutput TRUE for >= 5s continuous  | Held until 3s cooldown done | After 3s cooldown done AND heater would be OFF | Timer-driven, latch    | BOOLEAN            |
 * | SensorFault        | Temp < 0 OR Temp > 100              | N/A (implicit)      | When temp returns to valid range                        | Implicit               | BOOLEAN (derived)  |
 * | HeaterStatus       | HeaterOutput = TRUE                 | Same as HeaterOutput | Same as HeaterOutput                                   | Display only           | BOOLEAN            |
 * | CurrentTemperature | Always updated                      | Per scan            | N/A                                                     | Always active          | REAL, 0-100 valid  |
 *)

(* CONTRACT_RULES [{"kind":"hold_until_reset","output":"HeaterOutput","set_input":"OverheatProtection","reset_input":null}] *)

tmpSensorFault := (TemperatureSensorInput < 0.0) OR (TemperatureSensorInput > 100.0);

tmpHeaterShouldBeOn := (TemperatureSensorInput < SetTemperature) AND (NOT tmpSensorFault) AND (NOT OverheatProtection);

IF OverheatProtection THEN
    tonHeaterRuntime(IN := FALSE, PT := T#5S);
    tonOverheatCooldown(IN := TRUE, PT := T#3S);
    IF tonOverheatCooldown.Q THEN
        OverheatProtection := FALSE;
        tonOverheatCooldown(IN := FALSE, PT := T#3S);
    END_IF;
ELSIF tmpHeaterShouldBeOn THEN
    tonOverheatCooldown(IN := FALSE, PT := T#3S);
    tonHeaterRuntime(IN := TRUE, PT := T#5S);
    IF tonHeaterRuntime.Q THEN
        OverheatProtection := TRUE;
        HeaterOutput := FALSE;
    ELSE
        HeaterOutput := TRUE;
    END_IF;
ELSE
    tonHeaterRuntime(IN := FALSE, PT := T#5S);
    tonOverheatCooldown(IN := FALSE, PT := T#3S);
    HeaterOutput := FALSE;
END_IF;

CurrentTemperature := TemperatureSensorInput;
SetTempDisplay     := SetTemperature;
HeaterStatus       := HeaterOutput;

END_FUNCTION_BLOCK

(* ---- public-medium-04.raw_candidate_02.st ---- *)
FUNCTION_BLOCK FBTemperatureControl
VAR_INPUT
    TemperatureSensorInput : REAL;
    SetTemperature         : REAL;
END_VAR
VAR_OUTPUT
    CurrentTemperature : REAL;
    SetTempDisplay     : REAL;
    HeaterStatus       : BOOL;
    OverheatProtection : BOOL;
    HeaterOutput       : BOOL := FALSE;
END_VAR
VAR
    tonHeaterRuntime   : TON;
    tonOverheatCooldown: TON;
    tmpSensorFault     : BOOL;
END_VAR

(* ENGINEERING_CONTRACT:
 * | State/Output       | Activation                          | Retention           | Reset/Deactivation                                      | Same-scan Priority     | Units/Boundaries   |
 * |--------------------|-------------------------------------|---------------------|---------------------------------------------------------|------------------------|--------------------|
 * | HeaterOutput       | Temp < SetTemp AND no fault AND no overheat | Held per scan       | Temp >= SetTemp OR fault OR overheat triggered          | Overheat overrides     | BOOLEAN            |
 * | OverheatProtection | HeaterOutput TRUE for >= 5s continuous  | Held until 3s cooldown done | After 3s cooldown done AND heater would be OFF | Timer-driven, latch    | BOOLEAN            |
 * | SensorFault        | Temp < 0 OR Temp > 100              | N/A (implicit)      | When temp returns to valid range                        | Implicit               | BOOLEAN (derived)  |
 * | HeaterStatus       | HeaterOutput = TRUE                 | Same as HeaterOutput | Same as HeaterOutput                                   | Display only           | BOOLEAN            |
 * | CurrentTemperature | Always updated                      | Per scan            | N/A                                                     | Always active          | REAL, 0-100 valid  |
 *)

(* CONTRACT_RULES [] *)

tmpSensorFault := (TemperatureSensorInput < 0.0) OR (TemperatureSensorInput > 100.0);

IF OverheatProtection THEN
    tonHeaterRuntime(IN := FALSE, PT := T#0S);
    tonOverheatCooldown(IN := TRUE, PT := T#3S);
    IF tonOverheatCooldown.Q THEN
        OverheatProtection := FALSE;
        tonOverheatCooldown(IN := FALSE, PT := T#0S);
    END_IF;
    HeaterOutput := FALSE;
ELSIF (TemperatureSensorInput < SetTemperature) AND (NOT tmpSensorFault) THEN
    tonOverheatCooldown(IN := FALSE, PT := T#0S);
    tonHeaterRuntime(IN := TRUE, PT := T#5S);
    IF tonHeaterRuntime.Q THEN
        OverheatProtection := TRUE;
        HeaterOutput := FALSE;
        tonHeaterRuntime(IN := FALSE, PT := T#0S);
    ELSE
        HeaterOutput := TRUE;
    END_IF;
ELSE
    tonHeaterRuntime(IN := FALSE, PT := T#0S);
    tonOverheatCooldown(IN := FALSE, PT := T#0S);
    HeaterOutput := FALSE;
END_IF;

CurrentTemperature := TemperatureSensorInput;
SetTempDisplay     := SetTemperature;
HeaterStatus       := HeaterOutput;

END_FUNCTION_BLOCK

(* ---- public-medium-04.raw_candidate_03.st ---- *)
FUNCTION_BLOCK FBTemperatureControl
VAR_INPUT
    TemperatureSensorInput : REAL;
    SetTemperature         : REAL;
END_VAR
VAR_OUTPUT
    CurrentTemperature : REAL;
    SetTempDisplay     : REAL;
    HeaterStatus       : BOOL;
    OverheatProtection : BOOL;
    HeaterOutput       : BOOL := FALSE;
END_VAR
VAR
    tonOverheatCooldown : TON;
    tmpSensorFault      : BOOL;
    tmpHeaterShouldBeOn : BOOL;
    tmpHeaterOn         : BOOL;
    tmpRuntimeAccum     : LTIME;  // Track accumulated heating time
    tmpCooldownAccum    : LTIME;  // Track cooldown elapsed time
END_VAR

(* ENGINEERING_CONTRACT:
 * | State/Output       | Activation                          | Retention           | Reset/Deactivation                                      | Same-scan Priority     | Units/Boundaries   |
 * |--------------------|-------------------------------------|---------------------|---------------------------------------------------------|------------------------|--------------------|
 * | HeaterOutput       | Temp < SetTemp AND no fault AND no overheat | Held per scan   | Temp >= SetTemp OR fault OR overheat triggered          | Overheat overrides     | BOOLEAN            |
 * | OverheatProtection | Runtime >= 5s continuous heater ON  | Held until 3s cooldown done | After 3s cooldown done AND heater would be OFF | Timer-driven, latch    | BOOLEAN            |
 * | SensorFault        | Temp < 0 OR Temp > 100              | N/A (implicit)      | When temp returns to valid range                        | Implicit               | BOOLEAN (derived)  |
 * | HeaterStatus       | HeaterOutput = TRUE                 | Same as HeaterOutput | Same as HeaterOutput                                   | Display only           | BOOLEAN            |
 * | CurrentTemperature | Always updated                      | Per scan            | N/A                                                     | Always active          | REAL, 0-100 valid  |
 * | RuntimeAccum       | Increments when heater ON, no overheat | Per scan         | Reset when heater OFF OR overheat triggers             | Counter-based          | LTIME, max 5s      |
 * | CooldownAccum      | Increments when OverheatProtection TRUE | Per scan        | Reset when OverheatProtection clears                   | Counter-based          | LTIME, max 3s      |
 *)

(* CONTRACT_RULES [] *)

tmpSensorFault := (TemperatureSensorInput < 0.0) OR (TemperatureSensorInput > 100.0);

tmpHeaterOn := FALSE;

IF OverheatProtection THEN
    // Cooldown phase: heater stays off, track cooldown time
    tonOverheatCooldown(IN := TRUE, PT := T#3S);
    tmpCooldownAccum := tmpCooldownAccum + LTIME#1ms;  // Framework advances 1ms per call

    IF tonOverheatCooldown.Q THEN
        OverheatProtection := FALSE;
        tmpRuntimeAccum := LTIME#0ms;
        tonOverheatCooldown(IN := FALSE, PT := T#3S);
    END_IF;

ELSIF (NOT tmpSensorFault) AND (TemperatureSensorInput < SetTemperature) THEN
    // Normal heating: heater can be ON
    tonOverheatCooldown(IN := FALSE, PT := T#3S);

    tmpRuntimeAccum := tmpRuntimeAccum + LTIME#1ms;  // Framework advances 1ms per call

    IF tmpRuntimeAccum >= LTIME#5000ms THEN
        // Overheat threshold reached
        OverheatProtection := TRUE;
        HeaterOutput       := FALSE;
        tmpHeaterOn        := FALSE;
        tmpCooldownAccum   := LTIME#0ms;
    ELSE
        HeaterOutput := TRUE;
        tmpHeaterOn  := TRUE;
    END_IF;

ELSE
    // Temperature OK or sensor fault: heater OFF
    tonOverheatCooldown(IN := FALSE, PT := T#3S);
    HeaterOutput    := FALSE;
    tmpHeaterOn     := FALSE;
    tmpRuntimeAccum := LTIME#0ms;
END_IF;

CurrentTemperature := TemperatureSensorInput;
SetTempDisplay     := SetTemperature;
HeaterStatus       := tmpHeaterOn;

END_FUNCTION_BLOCK

(* ---- public-medium-04.raw_candidate_04.st ---- *)
FUNCTION_BLOCK FBTemperatureControl
VAR_INPUT
    TemperatureSensorInput : REAL;
    SetTemperature         : REAL;
END_VAR
VAR_OUTPUT
    CurrentTemperature : REAL;
    SetTempDisplay     : REAL;
    HeaterStatus       : BOOL;
    OverheatProtection : BOOL := FALSE;
    HeaterOutput       : BOOL := FALSE;
END_VAR
VAR
    tonHeaterRuntime   : TON;
    tonOverheatCooldown: TON;
    tmpSensorFault     : BOOL;
    tmpHeaterShouldBeOn: BOOL;
    tmpHeaterLatchedOff: BOOL := FALSE;
END_VAR

(* ENGINEERING_CONTRACT:
 * | State/Output       | Activation                          | Retention           | Reset/Deactivation                                      | Same-scan Priority     | Units/Boundaries   |
 * |--------------------|-------------------------------------|---------------------|---------------------------------------------------------|------------------------|--------------------|
 * | HeaterOutput       | Temp < SetTemp AND no fault AND no overheat/latch | Held per scan       | Temp >= SetTemp OR fault OR overheat/latch triggered    | Overheat overrides     | BOOLEAN            |
 * | OverheatProtection | HeaterOutput TRUE for >= 5s continuous  | Held until 3s cooldown done | After 3s cooldown done AND heater would be OFF | Timer-driven, latch    | BOOLEAN            |
 * | HeaterLatchedOff   | OverheatProtection triggers          | Held indefinitely   | No reset defined; remains latched                       | Latch persists         | BOOLEAN            |
 * | SensorFault        | Temp < 0 OR Temp > 100              | N/A (implicit)      | When temp returns to valid range                        | Implicit               | BOOLEAN (derived)  |
 * | HeaterStatus       | HeaterOutput = TRUE                 | Same as HeaterOutput | Same as HeaterOutput                                   | Display only           | BOOLEAN            |
 * | CurrentTemperature | Always updated                      | Per scan            | N/A                                                     | Always active          | REAL, 0-100 valid  |
 *)

(* CONTRACT_RULES [{"kind":"hold_until_reset","output":"HeaterOutput","set_input":"OverheatProtection","reset_input":null}] *)

tmpSensorFault := (TemperatureSensorInput < 0.0) OR (TemperatureSensorInput > 100.0);

IF OverheatProtection THEN
    tonHeaterRuntime(IN := FALSE, PT := T#5S);
    tonOverheatCooldown(IN := TRUE, PT := T#3S);
    IF tonOverheatCooldown.Q THEN
        OverheatProtection := FALSE;
        tmpHeaterLatchedOff := TRUE;
        tonOverheatCooldown(IN := FALSE, PT := T#3S);
        tonHeaterRuntime(IN := FALSE, PT := T#5S);
    END_IF;
    HeaterOutput := FALSE;
ELSIF tmpSensorFault THEN
    tonHeaterRuntime(IN := FALSE, PT := T#5S);
    tonOverheatCooldown(IN := FALSE, PT := T#3S);
    HeaterOutput := FALSE;
    tmpHeaterLatchedOff := FALSE;
ELSE
    tonOverheatCooldown(IN := FALSE, PT := T#3S);
    tmpHeaterShouldBeOn := (TemperatureSensorInput < SetTemperature) AND (NOT tmpHeaterLatchedOff);
    tonHeaterRuntime(IN := tmpHeaterShouldBeOn, PT := T#5S);
    IF tonHeaterRuntime.Q THEN
        OverheatProtection := TRUE;
        tmpHeaterLatchedOff := TRUE;
        HeaterOutput := FALSE;
    ELSIF tmpHeaterShouldBeOn THEN
        HeaterOutput := TRUE;
    ELSE
        HeaterOutput := FALSE;
        tmpHeaterLatchedOff := FALSE;
    END_IF;
END_IF;

CurrentTemperature := TemperatureSensorInput;
SetTempDisplay     := SetTemperature;
HeaterStatus       := HeaterOutput;

END_FUNCTION_BLOCK

(* ---- public-medium-08.candidate_01.st ---- *)
FUNCTION_BLOCK IPv4Parser
VAR_INPUT
    ipText : STRING(254);
END_VAR
VAR_OUTPUT
    ipValue : UDINT := 0;
END_VAR
VAR
    tmp_pos1      : INT;
    tmp_pos2      : INT;
    tmp_pos3      : INT;
    tmp_seg1      : STRING(4);
    tmp_seg2      : STRING(4);
    tmp_seg3      : STRING(4);
    tmp_seg4      : STRING(4);
    tmp_val1      : UDINT;
    tmp_val2      : UDINT;
    tmp_val3      : UDINT;
    tmp_val4      : UDINT;
    tmp_valid     : BOOL;
    tmp_i         : INT;
    tmp_char      : BYTE;
END_VAR
(* ENGINEERING_CONTRACT
  | Clause  | Output/State         | Behavior                                        |
  |---------|----------------------|-------------------------------------------------|
  | PUB001  | ipValue              | 32-bit UDINT; zero-initialized; updated once   |
  | PUB002  | ipValue              | RETENTION: holds last computed value           |
  | PUB002  | Validation path      | 4 segments via 3 period delimiters required    |
  | PUB003  | ipValue assembly     | Network byte order: seg1<<24 | seg2<<16 |      |
  |         |                      | seg3<<8 | seg4; SHL used for all shifts           |
  | PUB004  | Error output (0)     | SET: malformed, non-digit, count≠4, >255,      |
  |         |                      | or empty segment; RESET: none (latch to 0)     |
  | PUB004  | 0.0.0.0              | Produces 0; indistinguishable from error        |
  | General | Same-scan timing     | All segment extractions before any validation  |
  | General | Boundary: seg len    | 1-3 chars; non-digit check per character       |
  | General | Boundary: positions  | Periods must not be at index 0 or LEN-1        |
  | General | Type: LTIME/others   | Not applicable to this function block          |
  CONTRACT_RULES [] *)
BEGIN
    tmp_valid := TRUE;
    ipValue   := 0;

    tmp_pos1 := FIND(ipText, '.');
    tmp_pos2 := FIND(ipText, '.', tmp_pos1 + 1);
    tmp_pos3 := FIND(ipText, '.', tmp_pos2 + 1);

    tmp_valid := (tmp_pos1 > 0) AND (tmp_pos2 > tmp_pos1 + 1) AND (tmp_pos3 > tmp_pos2 + 1) AND (tmp_pos3 < LEN(ipText));

    IF tmp_valid THEN
        tmp_seg1 := MID(ipText, tmp_pos1 - 1, 1);
        tmp_seg2 := MID(ipText, tmp_pos2 - tmp_pos1 - 1, tmp_pos1 + 1);
        tmp_seg3 := MID(ipText, tmp_pos3 - tmp_pos2 - 1, tmp_pos2 + 1);
        tmp_seg4 := MID(ipText, LEN(ipText) - tmp_pos3, tmp_pos3 + 1);
    END_IF;

    IF tmp_valid THEN
        tmp_valid := (LEN(tmp_seg1) > 0) AND (LEN(tmp_seg2) > 0) AND (LEN(tmp_seg3) > 0) AND (LEN(tmp_seg4) > 0);
    END_IF;

    IF tmp_valid THEN
        FOR tmp_i := 1 TO LEN(tmp_seg1) DO
            tmp_char := tmp_seg1[tmp_i - 1];
            IF (tmp_char < 48) OR (tmp_char > 57) THEN
                tmp_valid := FALSE;
            END_IF;
        END_FOR;
    END_IF;

    IF tmp_valid THEN
        FOR tmp_i := 1 TO LEN(tmp_seg2) DO
            tmp_char := tmp_seg2[tmp_i - 1];
            IF (tmp_char < 48) OR (tmp_char > 57) THEN
                tmp_valid := FALSE;
            END_IF;
        END_FOR;
    END_IF;

    IF tmp_valid THEN
        FOR tmp_i := 1 TO LEN(tmp_seg3) DO
            tmp_char := tmp_seg3[tmp_i - 1];
            IF (tmp_char < 48) OR (tmp_char > 57) THEN
                tmp_valid := FALSE;
            END_IF;
        END_FOR;
    END_IF;

    IF tmp_valid THEN
        FOR tmp_i := 1 TO LEN(tmp_seg4) DO
            tmp_char := tmp_seg4[tmp_i - 1];
            IF (tmp_char < 48) OR (tmp_char > 57) THEN
                tmp_valid := FALSE;
            END_IF;
        END_FOR;
    END_IF;

    IF tmp_valid THEN
        tmp_val1 := TO_UDINT(TO_STRING(tmp_seg1));
        tmp_val2 := TO_UDINT(TO_STRING(tmp_seg2));
        tmp_val3 := TO_UDINT(TO_STRING(tmp_seg3));
        tmp_val4 := TO_UDINT(TO_STRING(tmp_seg4));

        tmp_valid := (tmp_val1 <= 255) AND (tmp_val2 <= 255) AND (tmp_val3 <= 255) AND (tmp_val4 <= 255);
    END_IF;

    IF tmp_valid THEN
        ipValue := SHL(tmp_val1, 24) OR SHL(tmp_val2, 16) OR SHL(tmp_val3, 8) OR tmp_val4;
    END_IF;
END_FUNCTION_BLOCK

(* ---- public-medium-08.candidate_02.st ---- *)
FUNCTION_BLOCK IPv4Parser
VAR_INPUT
    ipText : STRING(254);
END_VAR
VAR_OUTPUT
    ipValue : UDINT := 0;
END_VAR
VAR
    tmp_pos1      : INT;
    tmp_pos2      : INT;
    tmp_pos3      : INT;
    tmp_seg1      : STRING(4);
    tmp_seg2      : STRING(4);
    tmp_seg3      : STRING(4);
    tmp_seg4      : STRING(4);
    tmp_val1      : UDINT;
    tmp_val2      : UDINT;
    tmp_val3      : UDINT;
    tmp_val4      : UDINT;
    tmp_valid     : BOOL;
    tmp_i         : INT;
    tmp_char      : BYTE;
END_VAR
(* ENGINEERING_CONTRACT
  | Clause  | Output/State         | Behavior                                        |
  |---------|----------------------|-------------------------------------------------|
  | PUB001  | ipValue              | 32-bit UDINT; zero-initialized; updated once   |
  | PUB002  | ipValue              | RETENTION: holds last computed value           |
  | PUB002  | Validation path      | 4 segments via 3 period delimiters required    |
  | PUB003  | ipValue assembly     | Network byte order: seg1<<24 | seg2<<16 |      |
  |         |                      | seg3<<8 | seg4; SHL used for all shifts           |
  | PUB004  | Error output (0)     | SET: malformed, non-digit, count≠4, >255,      |
  |         |                      | or empty segment; RESET: none (latch to 0)     |
  | PUB004  | 0.0.0.0              | Produces 0; indistinguishable from error        |
  | General | Same-scan timing     | All segment extractions before any validation  |
  | General | Boundary: seg len    | 1-3 chars; non-digit check per character       |
  | General | Boundary: positions  | Periods must not be at index 0 or LEN-1        |
  | General | Type: LTIME/others   | Not applicable to this function block          |
  CONTRACT_RULES [] *)
BEGIN
    tmp_valid := TRUE;
    ipValue   := 0;

    tmp_pos1 := FIND(ipText, '.');
    tmp_pos2 := FIND(ipText, '.', tmp_pos1 + 1);
    tmp_pos3 := FIND(ipText, '.', tmp_pos2 + 1);

    tmp_valid := (tmp_pos1 > 0) AND (tmp_pos2 > tmp_pos1 + 1) AND (tmp_pos3 > tmp_pos2 + 1) AND (tmp_pos3 < LEN(ipText));

    IF tmp_valid THEN
        tmp_seg1 := MID(ipText, tmp_pos1 - 1, 1);
        tmp_seg2 := MID(ipText, tmp_pos2 - tmp_pos1 - 1, tmp_pos1 + 1);
        tmp_seg3 := MID(ipText, tmp_pos3 - tmp_pos2 - 1, tmp_pos2 + 1);
        tmp_seg4 := MID(ipText, LEN(ipText) - tmp_pos3, tmp_pos3 + 1);
    END_IF;

    IF tmp_valid THEN
        tmp_valid := (LEN(tmp_seg1) > 0) AND (LEN(tmp_seg2) > 0) AND (LEN(tmp_seg3) > 0) AND (LEN(tmp_seg4) > 0);
    END_IF;

    IF tmp_valid THEN
        FOR tmp_i := 1 TO LEN(tmp_seg1) DO
            tmp_char := tmp_seg1[tmp_i - 1];
            IF (tmp_char < 48) OR (tmp_char > 57) THEN
                tmp_valid := FALSE;
            END_IF;
        END_FOR;
    END_IF;

    IF tmp_valid THEN
        FOR tmp_i := 1 TO LEN(tmp_seg2) DO
            tmp_char := tmp_seg2[tmp_i - 1];
            IF (tmp_char < 48) OR (tmp_char > 57) THEN
                tmp_valid := FALSE;
            END_IF;
        END_FOR;
    END_IF;

    IF tmp_valid THEN
        FOR tmp_i := 1 TO LEN(tmp_seg3) DO
            tmp_char := tmp_seg3[tmp_i - 1];
            IF (tmp_char < 48) OR (tmp_char > 57) THEN
                tmp_valid := FALSE;
            END_IF;
        END_FOR;
    END_IF;

    IF tmp_valid THEN
        FOR tmp_i := 1 TO LEN(tmp_seg4) DO
            tmp_char := tmp_seg4[tmp_i - 1];
            IF (tmp_char < 48) OR (tmp_char > 57) THEN
                tmp_valid := FALSE;
            END_IF;
        END_FOR;
    END_IF;

    IF tmp_valid THEN
        tmp_val1 := TO_UDINT(tmp_seg1);
        tmp_val2 := TO_UDINT(tmp_seg2);
        tmp_val3 := TO_UDINT(tmp_seg3);
        tmp_val4 := TO_UDINT(tmp_seg4);

        tmp_valid := (tmp_val1 <= 255) AND (tmp_val2 <= 255) AND (tmp_val3 <= 255) AND (tmp_val4 <= 255);
    END_IF;

    IF tmp_valid THEN
        ipValue := SHL(tmp_val1, 24) OR SHL(tmp_val2, 16) OR SHL(tmp_val3, 8) OR tmp_val4;
    END_IF;
END_FUNCTION_BLOCK

(* ---- public-medium-08.candidate_03.st ---- *)
FUNCTION_BLOCK IPv4Parser
VAR_INPUT
    ipText : STRING(254);
END_VAR
VAR_OUTPUT
    ipValue : UDINT := 0;
END_VAR
VAR
    tmp_pos1      : INT;
    tmp_pos2      : INT;
    tmp_pos3      : INT;
    tmp_seg1      : STRING(4);
    tmp_seg2      : STRING(4);
    tmp_seg3      : STRING(4);
    tmp_seg4      : STRING(4);
    tmp_val1      : UDINT;
    tmp_val2      : UDINT;
    tmp_val3      : UDINT;
    tmp_val4      : UDINT;
    tmp_valid     : BOOL;
    tmp_i         : INT;
    tmp_char      : BYTE;
END_VAR
(* ENGINEERING_CONTRACT
  | Clause  | Output/State         | Behavior                                        |
  |---------|----------------------|-------------------------------------------------|
  | PUB001  | ipValue              | 32-bit UDINT; zero-initialized; updated once   |
  | PUB002  | ipValue              | RETENTION: holds last computed value           |
  | PUB002  | Validation path      | 4 segments via 3 period delimiters required    |
  | PUB003  | ipValue assembly     | Network byte order: seg1<<24 | seg2<<16 |      |
  |         |                      | seg3<<8 | seg4; SHL used for all shifts           |
  | PUB004  | Error output (0)     | SET: malformed, non-digit, count≠4, >255,      |
  |         |                      | or empty segment; RESET: none (latch to 0)     |
  | PUB004  | 0.0.0.0              | Produces 0; indistinguishable from error        |
  | General | Same-scan timing     | All segment extractions before any validation  |
  | General | Boundary: seg len    | 1-3 chars; non-digit check per character       |
  | General | Boundary: positions  | Periods must not be at index 0 or LEN-1        |
  | General | Type: LTIME/others   | Not applicable to this function block          |
  CONTRACT_RULES [] *)
BEGIN
    tmp_valid := TRUE;
    ipValue := 0;

    tmp_pos1 := FIND(ipText, '.');
    tmp_pos2 := FIND(ipText, '.', tmp_pos1 + 1);
    tmp_pos3 := FIND(ipText, '.', tmp_pos2 + 1);

    tmp_valid := (tmp_pos1 > 0) AND (tmp_pos2 > tmp_pos1 + 1) AND (tmp_pos3 > tmp_pos2 + 1) AND (tmp_pos3 < LEN(ipText));

    IF tmp_valid THEN
        tmp_seg1 := MID(ipText, tmp_pos1 - 1, 1);
        tmp_seg2 := MID(ipText, tmp_pos2 - tmp_pos1 - 1, tmp_pos1 + 1);
        tmp_seg3 := MID(ipText, tmp_pos3 - tmp_pos2 - 1, tmp_pos2 + 1);
        tmp_seg4 := MID(ipText, LEN(ipText) - tmp_pos3, tmp_pos3 + 1);
    END_IF;

    IF tmp_valid THEN
        tmp_valid := (LEN(tmp_seg1) > 0) AND (LEN(tmp_seg2) > 0) AND (LEN(tmp_seg3) > 0) AND (LEN(tmp_seg4) > 0);
    END_IF;

    IF tmp_valid THEN
        FOR tmp_i := 1 TO LEN(tmp_seg1) DO
            tmp_char := tmp_seg1[tmp_i - 1];
            IF (tmp_char < 48) OR (tmp_char > 57) THEN
                tmp_valid := FALSE;
            END_IF;
        END_FOR;
    END_IF;

    IF tmp_valid THEN
        FOR tmp_i := 1 TO LEN(tmp_seg2) DO
            tmp_char := tmp_seg2[tmp_i - 1];
            IF (tmp_char < 48) OR (tmp_char > 57) THEN
                tmp_valid := FALSE;
            END_IF;
        END_FOR;
    END_IF;

    IF tmp_valid THEN
        FOR tmp_i := 1 TO LEN(tmp_seg3) DO
            tmp_char := tmp_seg3[tmp_i - 1];
            IF (tmp_char < 48) OR (tmp_char > 57) THEN
                tmp_valid := FALSE;
            END_IF;
        END_FOR;
    END_IF;

    IF tmp_valid THEN
        FOR tmp_i := 1 TO LEN(tmp_seg4) DO
            tmp_char := tmp_seg4[tmp_i - 1];
            IF (tmp_char < 48) OR (tmp_char > 57) THEN
                tmp_valid := FALSE;
            END_IF;
        END_FOR;
    END_IF;

    IF tmp_valid THEN
        tmp_val1 := STRING_TO_UDINT(tmp_seg1);
        tmp_val2 := STRING_TO_UDINT(tmp_seg2);
        tmp_val3 := STRING_TO_UDINT(tmp_seg3);
        tmp_val4 := STRING_TO_UDINT(tmp_seg4);
        tmp_valid := (tmp_val1 <= 255) AND (tmp_val2 <= 255) AND (tmp_val3 <= 255) AND (tmp_val4 <= 255);
    END_IF;

    IF tmp_valid THEN
        ipValue := SHL(tmp_val1, 24) OR SHL(tmp_val2, 16) OR SHL(tmp_val3, 8) OR tmp_val4;
    END_IF;
END_FUNCTION_BLOCK

(* ---- public-medium-08.candidate_04.st ---- *)
FUNCTION_BLOCK IPv4Parser
VAR_INPUT
    ipText : STRING(254);
END_VAR
VAR_OUTPUT
    ipValue : UDINT := 0;
END_VAR
VAR
    tmp_pos1      : INT;
    tmp_pos2      : INT;
    tmp_pos3      : INT;
    tmp_seg1      : STRING(4);
    tmp_seg2      : STRING(4);
    tmp_seg3      : STRING(4);
    tmp_seg4      : STRING(4);
    tmp_val1      : UDINT;
    tmp_val2      : UDINT;
    tmp_val3      : UDINT;
    tmp_val4      : UDINT;
    tmp_valid     : BOOL;
    tmp_i         : INT;
    tmp_char      : BYTE;
    tmp_numeric   : BOOL;
END_VAR
(* ENGINEERING_CONTRACT
  | Clause  | Output/State         | Behavior                                        |
  |---------|----------------------|-------------------------------------------------|
  | PUB001  | ipValue              | 32-bit UDINT; zero-initialized; updated once   |
  | PUB002  | ipValue              | RETENTION: holds last computed value           |
  | PUB002  | Validation path      | 4 segments via 3 period delimiters required    |
  | PUB003  | ipValue assembly     | Network byte order: seg1<<24 | seg2<<16 |      |
  |         |                      | seg3<<8 | seg4; SHL used for all shifts           |
  | PUB004  | Error output (0)     | SET: malformed, non-digit, count≠4, >255,      |
  |         |                      | or empty segment; RESET: none (latch to 0)     |
  | PUB004  | 0.0.0.0              | Produces 0; indistinguishable from error        |
  | General | Same-scan timing     | All segment extractions before any validation  |
  | General | Boundary: seg len    | 1-3 chars; non-digit check per character       |
  | General | Boundary: positions  | Periods must not be at index 0 or LEN-1        |
  CONTRACT_RULES [] *)
BEGIN
    tmp_valid := TRUE;
    ipValue := 0;

    tmp_pos1 := FIND(ipText, '.');
    tmp_pos2 := FIND(ipText, '.', tmp_pos1 + 1);
    tmp_pos3 := FIND(ipText, '.', tmp_pos2 + 1);

    tmp_valid := (tmp_pos1 > 0) AND (tmp_pos2 > tmp_pos1 + 1) AND (tmp_pos3 > tmp_pos2 + 1) AND (tmp_pos3 < LEN(ipText));

    IF tmp_valid THEN
        tmp_seg1 := MID(ipText, tmp_pos1 - 1, 1);
        tmp_seg2 := MID(ipText, tmp_pos2 - tmp_pos1 - 1, tmp_pos1 + 1);
        tmp_seg3 := MID(ipText, tmp_pos3 - tmp_pos2 - 1, tmp_pos2 + 1);
        tmp_seg4 := MID(ipText, LEN(ipText) - tmp_pos3, tmp_pos3 + 1);
    END_IF;

    IF tmp_valid THEN
        tmp_valid := (LEN(tmp_seg1) >= 1) AND (LEN(tmp_seg1) <= 3) AND
                     (LEN(tmp_seg2) >= 1) AND (LEN(tmp_seg2) <= 3) AND
                     (LEN(tmp_seg3) >= 1) AND (LEN(tmp_seg3) <= 3) AND
                     (LEN(tmp_seg4) >= 1) AND (LEN(tmp_seg4) <= 3);
    END_IF;

    IF tmp_valid THEN
        FOR tmp_i := 0 TO LEN(tmp_seg1) - 1 DO
            tmp_char := tmp_seg1[tmp_i];
            tmp_numeric := (tmp_char >= 48) AND (tmp_char <= 57);
            IF NOT tmp_numeric THEN
                tmp_valid := FALSE;
            END_IF;
        END_FOR;
    END_IF;

    IF tmp_valid THEN
        FOR tmp_i := 0 TO LEN(tmp_seg2) - 1 DO
            tmp_char := tmp_seg2[tmp_i];
            tmp_numeric := (tmp_char >= 48) AND (tmp_char <= 57);
            IF NOT tmp_numeric THEN
                tmp_valid := FALSE;
            END_IF;
        END_FOR;
    END_IF;

    IF tmp_valid THEN
        FOR tmp_i := 0 TO LEN(tmp_seg3) - 1 DO
            tmp_char := tmp_seg3[tmp_i];
            tmp_numeric := (tmp_char >= 48) AND (tmp_char <= 57);
            IF NOT tmp_numeric THEN
                tmp_valid := FALSE;
            END_IF;
        END_FOR;
    END_IF;

    IF tmp_valid THEN
        FOR tmp_i := 0 TO LEN(tmp_seg4) - 1 DO
            tmp_char := tmp_seg4[tmp_i];
            tmp_numeric := (tmp_char >= 48) AND (tmp_char <= 57);
            IF NOT tmp_numeric THEN
                tmp_valid := FALSE;
            END_IF;
        END_FOR;
    END_IF;

    IF tmp_valid THEN
        tmp_val1 := TO_UDINT(tmp_seg1);
        tmp_val2 := TO_UDINT(tmp_seg2);
        tmp_val3 := TO_UDINT(tmp_seg3);
        tmp_val4 := TO_UDINT(tmp_seg4);

        tmp_valid := (tmp_val1 <= 255) AND (tmp_val2 <= 255) AND (tmp_val3 <= 255) AND (tmp_val4 <= 255);
    END_IF;

    IF tmp_valid THEN
        ipValue := SHL(tmp_val1, 24) OR SHL(tmp_val2, 16) OR SHL(tmp_val3, 8) OR tmp_val4;
    END_IF;
END_FUNCTION_BLOCK

(* ---- public-medium-08.raw_candidate_01.st ---- *)
FUNCTION_BLOCK IPv4Parser
VAR_INPUT
    ipText : STRING(254);
END_VAR
VAR_OUTPUT
    ipValue : UDINT := 0;
END_VAR
VAR
    tmp_pos1      : INT;
    tmp_pos2      : INT;
    tmp_pos3      : INT;
    tmp_seg1      : STRING(4);
    tmp_seg2      : STRING(4);
    tmp_seg3      : STRING(4);
    tmp_seg4      : STRING(4);
    tmp_val1      : UDINT;
    tmp_val2      : UDINT;
    tmp_val3      : UDINT;
    tmp_val4      : UDINT;
    tmp_valid     : BOOL;
    tmp_i         : INT;
    tmp_char      : BYTE;
END_VAR
(* ENGINEERING_CONTRACT
  | Clause  | Output/State         | Behavior                                        |
  |---------|----------------------|-------------------------------------------------|
  | PUB001  | ipValue              | 32-bit UDINT; zero-initialized; updated once   |
  | PUB002  | ipValue              | RETENTION: holds last computed value           |
  | PUB002  | Validation path      | 4 segments via 3 period delimiters required    |
  | PUB003  | ipValue assembly     | Network byte order: seg1<<24 | seg2<<16 |      |
  |         |                      | seg3<<8 | seg4; SHL used for all shifts           |
  | PUB004  | Error output (0)     | SET: malformed, non-digit, count≠4, >255,      |
  |         |                      | or empty segment; RESET: none (latch to 0)     |
  | PUB004  | 0.0.0.0              | Produces 0; indistinguishable from error        |
  | General | Same-scan timing     | All segment extractions before any validation  |
  | General | Boundary: seg len    | 1-3 chars; non-digit check per character       |
  | General | Boundary: positions  | Periods must not be at index 0 or LEN-1        |
  | General | Type: LTIME/others   | Not applicable to this function block          |
  CONTRACT_RULES [] *)
BEGIN
    tmp_valid := TRUE;
    ipValue   := 0;

    tmp_pos1 := FIND(ipText, '.');
    tmp_pos2 := FIND(ipText, '.', tmp_pos1 + 1);
    tmp_pos3 := FIND(ipText, '.', tmp_pos2 + 1);

    tmp_valid := (tmp_pos1 > 0) AND (tmp_pos2 > tmp_pos1 + 1) AND (tmp_pos3 > tmp_pos2 + 1) AND (tmp_pos3 < LEN(ipText));

    IF tmp_valid THEN
        tmp_seg1 := MID(ipText, tmp_pos1 - 1, 1);
        tmp_seg2 := MID(ipText, tmp_pos2 - tmp_pos1 - 1, tmp_pos1 + 1);
        tmp_seg3 := MID(ipText, tmp_pos3 - tmp_pos2 - 1, tmp_pos2 + 1);
        tmp_seg4 := MID(ipText, LEN(ipText) - tmp_pos3, tmp_pos3 + 1);
    END_IF;

    IF tmp_valid THEN
        tmp_valid := (LEN(tmp_seg1) > 0) AND (LEN(tmp_seg2) > 0) AND (LEN(tmp_seg3) > 0) AND (LEN(tmp_seg4) > 0);
    END_IF;

    IF tmp_valid THEN
        FOR tmp_i := 1 TO LEN(tmp_seg1) DO
            tmp_char := tmp_seg1[tmp_i - 1];
            IF (tmp_char < 48) OR (tmp_char > 57) THEN
                tmp_valid := FALSE;
            END_IF;
        END_FOR;
    END_IF;

    IF tmp_valid THEN
        FOR tmp_i := 1 TO LEN(tmp_seg2) DO
            tmp_char := tmp_seg2[tmp_i - 1];
            IF (tmp_char < 48) OR (tmp_char > 57) THEN
                tmp_valid := FALSE;
            END_IF;
        END_FOR;
    END_IF;

    IF tmp_valid THEN
        FOR tmp_i := 1 TO LEN(tmp_seg3) DO
            tmp_char := tmp_seg3[tmp_i - 1];
            IF (tmp_char < 48) OR (tmp_char > 57) THEN
                tmp_valid := FALSE;
            END_IF;
        END_FOR;
    END_IF;

    IF tmp_valid THEN
        FOR tmp_i := 1 TO LEN(tmp_seg4) DO
            tmp_char := tmp_seg4[tmp_i - 1];
            IF (tmp_char < 48) OR (tmp_char > 57) THEN
                tmp_valid := FALSE;
            END_IF;
        END_FOR;
    END_IF;

    IF tmp_valid THEN
        tmp_val1 := TO_UDINT(TO_STRING(tmp_seg1));
        tmp_val2 := TO_UDINT(TO_STRING(tmp_seg2));
        tmp_val3 := TO_UDINT(TO_STRING(tmp_seg3));
        tmp_val4 := TO_UDINT(TO_STRING(tmp_seg4));

        tmp_valid := (tmp_val1 <= 255) AND (tmp_val2 <= 255) AND (tmp_val3 <= 255) AND (tmp_val4 <= 255);
    END_IF;

    IF tmp_valid THEN
        ipValue := SHL(tmp_val1, 24) OR SHL(tmp_val2, 16) OR SHL(tmp_val3, 8) OR tmp_val4;
    END_IF;
END_FUNCTION_BLOCK

(* ---- public-medium-08.raw_candidate_02.st ---- *)
FUNCTION_BLOCK IPv4Parser
VAR_INPUT
    ipText : STRING(254);
END_VAR
VAR_OUTPUT
    ipValue : UDINT := 0;
END_VAR
VAR
    tmp_pos1      : INT;
    tmp_pos2      : INT;
    tmp_pos3      : INT;
    tmp_seg1      : STRING(4);
    tmp_seg2      : STRING(4);
    tmp_seg3      : STRING(4);
    tmp_seg4      : STRING(4);
    tmp_val1      : UDINT;
    tmp_val2      : UDINT;
    tmp_val3      : UDINT;
    tmp_val4      : UDINT;
    tmp_valid     : BOOL;
    tmp_i         : INT;
    tmp_char      : BYTE;
END_VAR
(* ENGINEERING_CONTRACT
  | Clause  | Output/State         | Behavior                                        |
  |---------|----------------------|-------------------------------------------------|
  | PUB001  | ipValue              | 32-bit UDINT; zero-initialized; updated once   |
  | PUB002  | ipValue              | RETENTION: holds last computed value           |
  | PUB002  | Validation path      | 4 segments via 3 period delimiters required    |
  | PUB003  | ipValue assembly     | Network byte order: seg1<<24 | seg2<<16 |      |
  |         |                      | seg3<<8 | seg4; SHL used for all shifts           |
  | PUB004  | Error output (0)     | SET: malformed, non-digit, count≠4, >255,      |
  |         |                      | or empty segment; RESET: none (latch to 0)     |
  | PUB004  | 0.0.0.0              | Produces 0; indistinguishable from error        |
  | General | Same-scan timing     | All segment extractions before any validation  |
  | General | Boundary: seg len    | 1-3 chars; non-digit check per character       |
  | General | Boundary: positions  | Periods must not be at index 0 or LEN-1        |
  | General | Type: LTIME/others   | Not applicable to this function block          |
  CONTRACT_RULES [] *)
BEGIN
    tmp_valid := TRUE;
    ipValue   := 0;

    tmp_pos1 := FIND(ipText, '.');
    tmp_pos2 := FIND(ipText, '.', tmp_pos1 + 1);
    tmp_pos3 := FIND(ipText, '.', tmp_pos2 + 1);

    tmp_valid := (tmp_pos1 > 0) AND (tmp_pos2 > tmp_pos1 + 1) AND (tmp_pos3 > tmp_pos2 + 1) AND (tmp_pos3 < LEN(ipText));

    IF tmp_valid THEN
        tmp_seg1 := MID(ipText, tmp_pos1 - 1, 1);
        tmp_seg2 := MID(ipText, tmp_pos2 - tmp_pos1 - 1, tmp_pos1 + 1);
        tmp_seg3 := MID(ipText, tmp_pos3 - tmp_pos2 - 1, tmp_pos2 + 1);
        tmp_seg4 := MID(ipText, LEN(ipText) - tmp_pos3, tmp_pos3 + 1);
    END_IF;

    IF tmp_valid THEN
        tmp_valid := (LEN(tmp_seg1) > 0) AND (LEN(tmp_seg2) > 0) AND (LEN(tmp_seg3) > 0) AND (LEN(tmp_seg4) > 0);
    END_IF;

    IF tmp_valid THEN
        FOR tmp_i := 1 TO LEN(tmp_seg1) DO
            tmp_char := tmp_seg1[tmp_i - 1];
            IF (tmp_char < 48) OR (tmp_char > 57) THEN
                tmp_valid := FALSE;
            END_IF;
        END_FOR;
    END_IF;

    IF tmp_valid THEN
        FOR tmp_i := 1 TO LEN(tmp_seg2) DO
            tmp_char := tmp_seg2[tmp_i - 1];
            IF (tmp_char < 48) OR (tmp_char > 57) THEN
                tmp_valid := FALSE;
            END_IF;
        END_FOR;
    END_IF;

    IF tmp_valid THEN
        FOR tmp_i := 1 TO LEN(tmp_seg3) DO
            tmp_char := tmp_seg3[tmp_i - 1];
            IF (tmp_char < 48) OR (tmp_char > 57) THEN
                tmp_valid := FALSE;
            END_IF;
        END_FOR;
    END_IF;

    IF tmp_valid THEN
        FOR tmp_i := 1 TO LEN(tmp_seg4) DO
            tmp_char := tmp_seg4[tmp_i - 1];
            IF (tmp_char < 48) OR (tmp_char > 57) THEN
                tmp_valid := FALSE;
            END_IF;
        END_FOR;
    END_IF;

    IF tmp_valid THEN
        tmp_val1 := TO_UDINT(tmp_seg1);
        tmp_val2 := TO_UDINT(tmp_seg2);
        tmp_val3 := TO_UDINT(tmp_seg3);
        tmp_val4 := TO_UDINT(tmp_seg4);

        tmp_valid := (tmp_val1 <= 255) AND (tmp_val2 <= 255) AND (tmp_val3 <= 255) AND (tmp_val4 <= 255);
    END_IF;

    IF tmp_valid THEN
        ipValue := SHL(tmp_val1, 24) OR SHL(tmp_val2, 16) OR SHL(tmp_val3, 8) OR tmp_val4;
    END_IF;
END_FUNCTION_BLOCK

(* ---- public-medium-08.raw_candidate_03.st ---- *)
FUNCTION_BLOCK IPv4Parser
VAR_INPUT
    ipText : STRING(254);
END_VAR
VAR_OUTPUT
    ipValue : UDINT := 0;
END_VAR
VAR
    tmp_pos1      : INT;
    tmp_pos2      : INT;
    tmp_pos3      : INT;
    tmp_seg1      : STRING(4);
    tmp_seg2      : STRING(4);
    tmp_seg3      : STRING(4);
    tmp_seg4      : STRING(4);
    tmp_val1      : UDINT;
    tmp_val2      : UDINT;
    tmp_val3      : UDINT;
    tmp_val4      : UDINT;
    tmp_valid     : BOOL;
    tmp_i         : INT;
    tmp_char      : BYTE;
END_VAR
(* ENGINEERING_CONTRACT
  | Clause  | Output/State         | Behavior                                        |
  |---------|----------------------|-------------------------------------------------|
  | PUB001  | ipValue              | 32-bit UDINT; zero-initialized; updated once   |
  | PUB002  | ipValue              | RETENTION: holds last computed value           |
  | PUB002  | Validation path      | 4 segments via 3 period delimiters required    |
  | PUB003  | ipValue assembly     | Network byte order: seg1<<24 | seg2<<16 |      |
  |         |                      | seg3<<8 | seg4; SHL used for all shifts           |
  | PUB004  | Error output (0)     | SET: malformed, non-digit, count≠4, >255,      |
  |         |                      | or empty segment; RESET: none (latch to 0)     |
  | PUB004  | 0.0.0.0              | Produces 0; indistinguishable from error        |
  | General | Same-scan timing     | All segment extractions before any validation  |
  | General | Boundary: seg len    | 1-3 chars; non-digit check per character       |
  | General | Boundary: positions  | Periods must not be at index 0 or LEN-1        |
  | General | Type: LTIME/others   | Not applicable to this function block          |
  CONTRACT_RULES [] *)
BEGIN
    tmp_valid := TRUE;
    ipValue := 0;

    tmp_pos1 := FIND(ipText, '.');
    tmp_pos2 := FIND(ipText, '.', tmp_pos1 + 1);
    tmp_pos3 := FIND(ipText, '.', tmp_pos2 + 1);

    tmp_valid := (tmp_pos1 > 0) AND (tmp_pos2 > tmp_pos1 + 1) AND (tmp_pos3 > tmp_pos2 + 1) AND (tmp_pos3 < LEN(ipText));

    IF tmp_valid THEN
        tmp_seg1 := MID(ipText, tmp_pos1 - 1, 1);
        tmp_seg2 := MID(ipText, tmp_pos2 - tmp_pos1 - 1, tmp_pos1 + 1);
        tmp_seg3 := MID(ipText, tmp_pos3 - tmp_pos2 - 1, tmp_pos2 + 1);
        tmp_seg4 := MID(ipText, LEN(ipText) - tmp_pos3, tmp_pos3 + 1);
    END_IF

    IF tmp_valid THEN
        tmp_valid := (LEN(tmp_seg1) > 0) AND (LEN(tmp_seg2) > 0) AND (LEN(tmp_seg3) > 0) AND (LEN(tmp_seg4) > 0);
    END_IF

    IF tmp_valid THEN
        FOR tmp_i := 1 TO LEN(tmp_seg1) DO
            tmp_char := tmp_seg1[tmp_i - 1];
            IF (tmp_char < 48) OR (tmp_char > 57) THEN
                tmp_valid := FALSE;
            END_IF;
        END_FOR;
    END_IF

    IF tmp_valid THEN
        FOR tmp_i := 1 TO LEN(tmp_seg2) DO
            tmp_char := tmp_seg2[tmp_i - 1];
            IF (tmp_char < 48) OR (tmp_char > 57) THEN
                tmp_valid := FALSE;
            END_IF;
        END_FOR;
    END_IF

    IF tmp_valid THEN
        FOR tmp_i := 1 TO LEN(tmp_seg3) DO
            tmp_char := tmp_seg3[tmp_i - 1];
            IF (tmp_char < 48) OR (tmp_char > 57) THEN
                tmp_valid := FALSE;
            END_IF;
        END_FOR;
    END_IF

    IF tmp_valid THEN
        FOR tmp_i := 1 TO LEN(tmp_seg4) DO
            tmp_char := tmp_seg4[tmp_i - 1];
            IF (tmp_char < 48) OR (tmp_char > 57) THEN
                tmp_valid := FALSE;
            END_IF;
        END_FOR;
    END_IF

    IF tmp_valid THEN
        tmp_val1 := STRING_TO_UDINT(tmp_seg1);
        tmp_val2 := STRING_TO_UDINT(tmp_seg2);
        tmp_val3 := STRING_TO_UDINT(tmp_seg3);
        tmp_val4 := STRING_TO_UDINT(tmp_seg4);
        tmp_valid := (tmp_val1 <= 255) AND (tmp_val2 <= 255) AND (tmp_val3 <= 255) AND (tmp_val4 <= 255);
    END_IF

    IF tmp_valid THEN
        ipValue := SHL(tmp_val1, 24) OR SHL(tmp_val2, 16) OR SHL(tmp_val3, 8) OR tmp_val4;
    END_IF
END_FUNCTION_BLOCK
